//     Term 34 (AT2200-0500)/CC Inputs/Current actual value Ch.23 <-> Data Pointer/CurrentActualValues[22]
//     Term 34 (AT2200-0500)/CC Inputs/Current actual value Ch.24 <-> Data Pointer/CurrentActualValues[23]
//     Term 34 (AT2200-0500)/CC Inputs/Current actual value Ch.25 <-> Data Pointer/CurrentActualValues[24]
//     Term 34 (AT2200-0500)/CC Inputs/Current actual value Ch.26 <-> Data Pointer/CurrentActualValues[25]
//     Term 34 (AT2200-0500)/CC Inputs/Current actual value Ch.27 <-> Data Pointer/CurrentActualValues[26]
//     Term 34 (AT2200-0500)/CC Inputs/Current actual value Ch.28 <-> Data Pointer/CurrentActualValues[27]
//     Term 34 (AT2200-0500)/CC Inputs/Current actual value Ch.29 <-> Data Pointer/CurrentActualValues[28]
//     Term 34 (AT2200-0500)/CC Inputs/Current actual value Ch.3 <-> Data Pointer/CurrentActualValues[2]
//     Term 34 (AT2200-0500)/CC Inputs/Current actual value Ch.30 <-> Data Pointer/CurrentActualValues[29]
//     Term 34 (AT2200-0500)/CC Inputs/Current actual value Ch.4 <-> Data Pointer/CurrentActualValues[3]
//     Term 34 (AT2200-0500)/CC Inputs/Current actual value Ch.5 <-> Data Pointer/CurrentActualValues[4]
//     Term 34 (AT2200-0500)/CC Inputs/Current actual value Ch.6 <-> Data Pointer/CurrentActualValues[5]
//     Term 34 (AT2200-0500)/CC Inputs/Current actual value Ch.7 <-> Data Pointer/CurrentActualValues[6]
//     Term 34 (AT2200-0500)/CC Inputs/Current actual value Ch.8 <-> Data Pointer/CurrentActualValues[7]
//     Term 34 (AT2200-0500)/CC Inputs/Current actual value Ch.9 <-> Data Pointer/CurrentActualValues[8]
//     Term 34 (AT2200-0500)/CC Inputs/Status <-> Data Pointer/Status
//     Term 34 (AT2200-0500)/CC Outputs/Control <-> Data Pointer/Control
//     Term 34 (AT2200-0500)/CC Outputs/Current setpoint value Ch.1 <-> Data Pointer/CurrentSetpointValues[0]
//     Term 34 (AT2200-0500)/CC Outputs/Current setpoint value Ch.10 <-> Data Pointer/CurrentSetpointValues[9]
//     Term 34 (AT2200-0500)/CC Outputs/Current setpoint value Ch.11 <-> Data Pointer/CurrentSetpointValues[10]
//     Term 34 (AT2200-0500)/CC Outputs/Current setpoint value Ch.12 <-> Data Pointer/CurrentSetpointValues[11]
//     Term 34 (AT2200-0500)/CC Outputs/Current setpoint value Ch.13 <-> Data Pointer/CurrentSetpointValues[12]
//     Term 34 (AT2200-0500)/CC Outputs/Current setpoint value Ch.14 <-> Data Pointer/CurrentSetpointValues[13]
//     Term 34 (AT2200-0500)/CC Outputs/Current setpoint value Ch.15 <-> Data Pointer/CurrentSetpointValues[14]
//     Term 34 (AT2200-0500)/CC Outputs/Current setpoint value Ch.16 <-> Data Pointer/CurrentSetpointValues[15]
//     Term 34 (AT2200-0500)/CC Outputs/Current setpoint value Ch.17 <-> Data Pointer/CurrentSetpointValues[16]
//     Term 34 (AT2200-0500)/CC Outputs/Current setpoint value Ch.18 <-> Data Pointer/CurrentSetpointValues[17]
//     Term 34 (AT2200-0500)/CC Outputs/Current setpoint value Ch.19 <-> Data Pointer/CurrentSetpointValues[18]
//     Term 34 (AT2200-0500)/CC Outputs/Current setpoint value Ch.2 <-> Data Pointer/CurrentSetpointValues[1]
//     Term 34 (AT2200-0500)/CC Outputs/Current setpoint value Ch.20 <-> Data Pointer/CurrentSetpointValues[19]
//     Term 34 (AT2200-0500)/CC Outputs/Current setpoint value Ch.21 <-> Data Pointer/CurrentSetpointValues[20]
//     Term 34 (AT2200-0500)/CC Outputs/Current setpoint value Ch.22 <-> Data Pointer/CurrentSetpointValues[21]
//     Term 34 (AT2200-0500)/CC Outputs/Current setpoint value Ch.23 <-> Data Pointer/CurrentSetpointValues[22]
//     Term 34 (AT2200-0500)/CC Outputs/Current setpoint value Ch.24 <-> Data Pointer/CurrentSetpointValues[23]
//     Term 34 (AT2200-0500)/CC Outputs/Current setpoint value Ch.25 <-> Data Pointer/CurrentSetpointValues[24]
//     Term 34 (AT2200-0500)/CC Outputs/Current setpoint value Ch.26 <-> Data Pointer/CurrentSetpointValues[25]
//     Term 34 (AT2200-0500)/CC Outputs/Current setpoint value Ch.27 <-> Data Pointer/CurrentSetpointValues[26]
//     Term 34 (AT2200-0500)/CC Outputs/Current setpoint value Ch.28 <-> Data Pointer/CurrentSetpointValues[27]
//     Term 34 (AT2200-0500)/CC Outputs/Current setpoint value Ch.29 <-> Data Pointer/CurrentSetpointValues[28]
//     Term 34 (AT2200-0500)/CC Outputs/Current setpoint value Ch.3 <-> Data Pointer/CurrentSetpointValues[2]
//     Term 34 (AT2200-0500)/CC Outputs/Current setpoint value Ch.30 <-> Data Pointer/CurrentSetpointValues[29]
//     Term 34 (AT2200-0500)/CC Outputs/Current setpoint value Ch.4 <-> Data Pointer/CurrentSetpointValues[3]
//     Term 34 (AT2200-0500)/CC Outputs/Current setpoint value Ch.5 <-> Data Pointer/CurrentSetpointValues[4]
//     Term 34 (AT2200-0500)/CC Outputs/Current setpoint value Ch.6 <-> Data Pointer/CurrentSetpointValues[5]
//     Term 34 (AT2200-0500)/CC Outputs/Current setpoint value Ch.7 <-> Data Pointer/CurrentSetpointValues[6]
//     Term 34 (AT2200-0500)/CC Outputs/Current setpoint value Ch.8 <-> Data Pointer/CurrentSetpointValues[7]
//     Term 34 (AT2200-0500)/CC Outputs/Current setpoint value Ch.9 <-> Data Pointer/CurrentSetpointValues[8]
//     Term 34 (AT2200-0500)/LFB Inputs/BinaryData <-> Data Pointer/HallSensorValues
//   Device 36 <-> TcCOM Objects/XTS ProcessingUnit 1/Part 1/Module 42
//     Term 35 (AT2200-0500)/CC Inputs/Current actual value Ch.1 <-> Data Pointer/CurrentActualValues[0]
//     Term 35 (AT2200-0500)/CC Inputs/Current actual value Ch.10 <-> Data Pointer/CurrentActualValues[9]
//     Term 35 (AT2200-0500)/CC Inputs/Current actual value Ch.11 <-> Data Pointer/CurrentActualValues[10]
//     Term 35 (AT2200-0500)/CC Inputs/Current actual value Ch.12 <-> Data Pointer/CurrentActualValues[11]
//     Term 35 (AT2200-0500)/CC Inputs/Current actual value Ch.13 <-> Data Pointer/CurrentActualValues[12]
//     Term 35 (AT2200-0500)/CC Inputs/Current actual value Ch.14 <-> Data Pointer/CurrentActualValues[13]
//     Term 35 (AT2200-0500)/CC Inputs/Current actual value Ch.15 <-> Data Pointer/CurrentActualValues[14]
//     Term 35 (AT2200-0500)/CC Inputs/Current actual value Ch.16 <-> Data Pointer/CurrentActualValues[15]
//     Term 35 (AT2200-0500)/CC Inputs/Current actual value Ch.17 <-> Data Pointer/CurrentActualValues[16]
//     Term 35 (AT2200-0500)/CC Inputs/Current actual value Ch.18 <-> Data Pointer/CurrentActualValues[17]
//     Term 35 (AT2200-0500)/CC Inputs/Current actual value Ch.19 <-> Data Pointer/CurrentActualValues[18]
//     Term 35 (AT2200-0500)/CC Inputs/Current actual value Ch.2 <-> Data Pointer/CurrentActualValues[1]
//     Term 35 (AT2200-0500)/CC Inputs/Current actual value Ch.20 <-> Data Pointer/CurrentActualValues[19]
//     Term 35 (AT2200-0500)/CC Inputs/Current actual value Ch.21 <-> Data Pointer/CurrentActualValues[20]
//     Term 35 (AT2200-0500)/CC Inputs/Current actual value Ch.22 <-> Data Pointer/CurrentActualValues[21]
//     Term 35 (AT2200-0500)/CC Inputs/Current actual value Ch.23 <-> Data Pointer/CurrentActualValues[22]
//     Term 35 (AT2200-0500)/CC Inputs/Current actual value Ch.24 <-> Data Pointer/CurrentActualValues[23]
//     Term 35 (AT2200-0500)/CC Inputs/Current actual value Ch.25 <-> Data Pointer/CurrentActualValues[24]
//     Term 35 (AT2200-0500)/CC Inputs/Current actual value Ch.26 <-> Data Pointer/CurrentActualValues[25]
//     Term 35 (AT2200-0500)/CC Inputs/Current actual value Ch.27 <-> Data Pointer/CurrentActualValues[26]
//     Term 35 (AT2200-0500)/CC Inputs/Current actual value Ch.28 <-> Data Pointer/CurrentActualValues[27]
//     Term 35 (AT2200-0500)/CC Inputs/Current actual value Ch.29 <-> Data Pointer/CurrentActualValues[28]
//     Term 35 (AT2200-0500)/CC Inputs/Current actual value Ch.3 <-> Data Pointer/CurrentActualValues[2]
//     Term 35 (AT2200-0500)/CC Inputs/Current actual value Ch.30 <-> Data Pointer/CurrentActualValues[29]
//     Term 35 (AT2200-0500)/CC Inputs/Current actual value Ch.4 <-> Data Pointer/CurrentActualValues[3]
//     Term 35 (AT2200-0500)/CC Inputs/Current actual value Ch.5 <-> Data Pointer/CurrentActualValues[4]
//     Term 35 (AT2200-0500)/CC Inputs/Current actual value Ch.6 <-> Data Pointer/CurrentActualValues[5]
//     Term 35 (AT2200-0500)/CC Inputs/Current actual value Ch.7 <-> Data Pointer/CurrentActualValues[6]
//     Term 35 (AT2200-0500)/CC Inputs/Current actual value Ch.8 <-> Data Pointer/CurrentActualValues[7]
//     Term 35 (AT2200-0500)/CC Inputs/Current actual value Ch.9 <-> Data Pointer/CurrentActualValues[8]
//     Term 35 (AT2200-0500)/CC Inputs/Status <-> Data Pointer/Status
//     Term 35 (AT2200-0500)/CC Outputs/Control <-> Data Pointer/Control
//     Term 35 (AT2200-0500)/CC Outputs/Current setpoint value Ch.1 <-> Data Pointer/CurrentSetpointValues[0]
//     Term 35 (AT2200-0500)/CC Outputs/Current setpoint value Ch.10 <-> Data Pointer/CurrentSetpointValues[9]
//     Term 35 (AT2200-0500)/CC Outputs/Current setpoint value Ch.11 <-> Data Pointer/CurrentSetpointValues[10]
//     Term 35 (AT2200-0500)/CC Outputs/Current setpoint value Ch.12 <-> Data Pointer/CurrentSetpointValues[11]
//     Term 35 (AT2200-0500)/CC Outputs/Current setpoint value Ch.13 <-> Data Pointer/CurrentSetpointValues[12]
//     Term 35 (AT2200-0500)/CC Outputs/Current setpoint value Ch.14 <-> Data Pointer/CurrentSetpointValues[13]
//     Term 35 (AT2200-0500)/CC Outputs/Current setpoint value Ch.15 <-> Data Pointer/CurrentSetpointValues[14]
//     Term 35 (AT2200-0500)/CC Outputs/Current setpoint value Ch.16 <-> Data Pointer/CurrentSetpointValues[15]
//     Term 35 (AT2200-0500)/CC Outputs/Current setpoint value Ch.17 <-> Data Pointer/CurrentSetpointValues[16]
//     Term 35 (AT2200-0500)/CC Outputs/Current setpoint value Ch.18 <-> Data Pointer/CurrentSetpointValues[17]
//     Term 35 (AT2200-0500)/CC Outputs/Current setpoint value Ch.19 <-> Data Pointer/CurrentSetpointValues[18]
//     Term 35 (AT2200-0500)/CC Outputs/Current setpoint value Ch.2 <-> Data Pointer/CurrentSetpointValues[1]
//     Term 35 (AT2200-0500)/CC Outputs/Current setpoint value Ch.20 <-> Data Pointer/CurrentSetpointValues[19]
//     Term 35 (AT2200-0500)/CC Outputs/Current setpoint value Ch.21 <-> Data Pointer/CurrentSetpointValues[20]
//     Term 35 (AT2200-0500)/CC Outputs/Current setpoint value Ch.22 <-> Data Pointer/CurrentSetpointValues[21]
//     Term 35 (AT2200-0500)/CC Outputs/Current setpoint value Ch.23 <-> Data Pointer/CurrentSetpointValues[22]
//     Term 35 (AT2200-0500)/CC Outputs/Current setpoint value Ch.24 <-> Data Pointer/CurrentSetpointValues[23]
//     Term 35 (AT2200-0500)/CC Outputs/Current setpoint value Ch.25 <-> Data Pointer/CurrentSetpointValues[24]
//     Term 35 (AT2200-0500)/CC Outputs/Current setpoint value Ch.26 <-> Data Pointer/CurrentSetpointValues[25]
//     Term 35 (AT2200-0500)/CC Outputs/Current setpoint value Ch.27 <-> Data Pointer/CurrentSetpointValues[26]
//     Term 35 (AT2200-0500)/CC Outputs/Current setpoint value Ch.28 <-> Data Pointer/CurrentSetpointValues[27]
//     Term 35 (AT2200-0500)/CC Outputs/Current setpoint value Ch.29 <-> Data Pointer/CurrentSetpointValues[28]
//     Term 35 (AT2200-0500)/CC Outputs/Current setpoint value Ch.3 <-> Data Pointer/CurrentSetpointValues[2]
//     Term 35 (AT2200-0500)/CC Outputs/Current setpoint value Ch.30 <-> Data Pointer/CurrentSetpointValues[29]
//     Term 35 (AT2200-0500)/CC Outputs/Current setpoint value Ch.4 <-> Data Pointer/CurrentSetpointValues[3]
//     Term 35 (AT2200-0500)/CC Outputs/Current setpoint value Ch.5 <-> Data Pointer/CurrentSetpointValues[4]
//     Term 35 (AT2200-0500)/CC Outputs/Current setpoint value Ch.6 <-> Data Pointer/CurrentSetpointValues[5]
//     Term 35 (AT2200-0500)/CC Outputs/Current setpoint value Ch.7 <-> Data Pointer/CurrentSetpointValues[6]
//     Term 35 (AT2200-0500)/CC Outputs/Current setpoint value Ch.8 <-> Data Pointer/CurrentSetpointValues[7]
//     Term 35 (AT2200-0500)/CC Outputs/Current setpoint value Ch.9 <-> Data Pointer/CurrentSetpointValues[8]
//     Term 35 (AT2200-0500)/LFB Inputs/BinaryData <-> Data Pointer/HallSensorValues
//   Device 37 <-> TcCOM Objects/XTS ProcessingUnit 1/Part 1/Module 43
//     Term 36 (AT2202-0500)/CC Inputs/Current actual value Ch.1 <-> Data Pointer/CurrentActualValues[0]
//     Term 36 (AT2202-0500)/CC Inputs/Current actual value Ch.10 <-> Data Pointer/CurrentActualValues[9]
//     Term 36 (AT2202-0500)/CC Inputs/Current actual value Ch.11 <-> Data Pointer/CurrentActualValues[10]
//     Term 36 (AT2202-0500)/CC Inputs/Current actual value Ch.12 <-> Data Pointer/CurrentActualValues[11]
//     Term 36 (AT2202-0500)/CC Inputs/Current actual value Ch.13 <-> Data Pointer/CurrentActualValues[12]
//     Term 36 (AT2202-0500)/CC Inputs/Current actual value Ch.14 <-> Data Pointer/CurrentActualValues[13]
//     Term 36 (AT2202-0500)/CC Inputs/Current actual value Ch.15 <-> Data Pointer/CurrentActualValues[14]
//     Term 36 (AT2202-0500)/CC Inputs/Current actual value Ch.16 <-> Data Pointer/CurrentActualValues[15]
//     Term 36 (AT2202-0500)/CC Inputs/Current actual value Ch.17 <-> Data Pointer/CurrentActualValues[16]
//     Term 36 (AT2202-0500)/CC Inputs/Current actual value Ch.18 <-> Data Pointer/CurrentActualValues[17]
//     Term 36 (AT2202-0500)/CC Inputs/Current actual value Ch.19 <-> Data Pointer/CurrentActualValues[18]
//     Term 36 (AT2202-0500)/CC Inputs/Current actual value Ch.2 <-> Data Pointer/CurrentActualValues[1]
//     Term 36 (AT2202-0500)/CC Inputs/Current actual value Ch.20 <-> Data Pointer/CurrentActualValues[19]
//     Term 36 (AT2202-0500)/CC Inputs/Current actual value Ch.21 <-> Data Pointer/CurrentActualValues[20]
//     Term 36 (AT2202-0500)/CC Inputs/Current actual value Ch.22 <-> Data Pointer/CurrentActualValues[21]
//     Term 36 (AT2202-0500)/CC Inputs/Current actual value Ch.23 <-> Data Pointer/CurrentActualValues[22]
//     Term 36 (AT2202-0500)/CC Inputs/Current actual value Ch.24 <-> Data Pointer/CurrentActualValues[23]
//     Term 36 (AT2202-0500)/CC Inputs/Current actual value Ch.25 <-> Data Pointer/CurrentActualValues[24]
//     Term 36 (AT2202-0500)/CC Inputs/Current actual value Ch.26 <-> Data Pointer/CurrentActualValues[25]
//     Term 36 (AT2202-0500)/CC Inputs/Current actual value Ch.27 <-> Data Pointer/CurrentActualValues[26]
//     Term 36 (AT2202-0500)/CC Inputs/Current actual value Ch.28 <-> Data Pointer/CurrentActualValues[27]
//     Term 36 (AT2202-0500)/CC Inputs/Current actual value Ch.29 <-> Data Pointer/CurrentActualValues[28]
//     Term 36 (AT2202-0500)/CC Inputs/Current actual value Ch.3 <-> Data Pointer/CurrentActualValues[2]
//     Term 36 (AT2202-0500)/CC Inputs/Current actual value Ch.30 <-> Data Pointer/CurrentActualValues[29]
//     Term 36 (AT2202-0500)/CC Inputs/Current actual value Ch.4 <-> Data Pointer/CurrentActualValues[3]
//     Term 36 (AT2202-0500)/CC Inputs/Current actual value Ch.5 <-> Data Pointer/CurrentActualValues[4]
//     Term 36 (AT2202-0500)/CC Inputs/Current actual value Ch.6 <-> Data Pointer/CurrentActualValues[5]
//     Term 36 (AT2202-0500)/CC Inputs/Current actual value Ch.7 <-> Data Pointer/CurrentActualValues[6]
//     Term 36 (AT2202-0500)/CC Inputs/Current actual value Ch.8 <-> Data Pointer/CurrentActualValues[7]
//     Term 36 (AT2202-0500)/CC Inputs/Current actual value Ch.9 <-> Data Pointer/CurrentActualValues[8]
//     Term 36 (AT2202-0500)/CC Inputs/Status <-> Data Pointer/Status
//     Term 36 (AT2202-0500)/CC Outputs/Control <-> Data Pointer/Control
//     Term 36 (AT2202-0500)/CC Outputs/Current setpoint value Ch.1 <-> Data Pointer/CurrentSetpointValues[0]
//     Term 36 (AT2202-0500)/CC Outputs/Current setpoint value Ch.10 <-> Data Pointer/CurrentSetpointValues[9]
//     Term 36 (AT2202-0500)/CC Outputs/Current setpoint value Ch.11 <-> Data Pointer/CurrentSetpointValues[10]
//     Term 36 (AT2202-0500)/CC Outputs/Current setpoint value Ch.12 <-> Data Pointer/CurrentSetpointValues[11]
//     Term 36 (AT2202-0500)/CC Outputs/Current setpoint value Ch.13 <-> Data Pointer/CurrentSetpointValues[12]
//     Term 36 (AT2202-0500)/CC Outputs/Current setpoint value Ch.14 <-> Data Pointer/CurrentSetpointValues[13]
//     Term 36 (AT2202-0500)/CC Outputs/Current setpoint value Ch.15 <-> Data Pointer/CurrentSetpointValues[14]
//     Term 36 (AT2202-0500)/CC Outputs/Current setpoint value Ch.16 <-> Data Pointer/CurrentSetpointValues[15]
//     Term 36 (AT2202-0500)/CC Outputs/Current setpoint value Ch.17 <-> Data Pointer/CurrentSetpointValues[16]
//     Term 36 (AT2202-0500)/CC Outputs/Current setpoint value Ch.18 <-> Data Pointer/CurrentSetpointValues[17]
//     Term 36 (AT2202-0500)/CC Outputs/Current setpoint value Ch.19 <-> Data Pointer/CurrentSetpointValues[18]
//     Term 36 (AT2202-0500)/CC Outputs/Current setpoint value Ch.2 <-> Data Pointer/CurrentSetpointValues[1]
//     Term 36 (AT2202-0500)/CC Outputs/Current setpoint value Ch.20 <-> Data Pointer/CurrentSetpointValues[19]
//     Term 36 (AT2202-0500)/CC Outputs/Current setpoint value Ch.21 <-> Data Pointer/CurrentSetpointValues[20]
//     Term 36 (AT2202-0500)/CC Outputs/Current setpoint value Ch.22 <-> Data Pointer/CurrentSetpointValues[21]
//     Term 36 (AT2202-0500)/CC Outputs/Current setpoint value Ch.23 <-> Data Pointer/CurrentSetpointValues[22]
//     Term 36 (AT2202-0500)/CC Outputs/Current setpoint value Ch.24 <-> Data Pointer/CurrentSetpointValues[23]
//     Term 36 (AT2202-0500)/CC Outputs/Current setpoint value Ch.25 <-> Data Pointer/CurrentSetpointValues[24]
//     Term 36 (AT2202-0500)/CC Outputs/Current setpoint value Ch.26 <-> Data Pointer/CurrentSetpointValues[25]
//     Term 36 (AT2202-0500)/CC Outputs/Current setpoint value Ch.27 <-> Data Pointer/CurrentSetpointValues[26]
//     Term 36 (AT2202-0500)/CC Outputs/Current setpoint value Ch.28 <-> Data Pointer/CurrentSetpointValues[27]
//     Term 36 (AT2202-0500)/CC Outputs/Current setpoint value Ch.29 <-> Data Pointer/CurrentSetpointValues[28]
//     Term 36 (AT2202-0500)/CC Outputs/Current setpoint value Ch.3 <-> Data Pointer/CurrentSetpointValues[2]
//     Term 36 (AT2202-0500)/CC Outputs/Current setpoint value Ch.30 <-> Data Pointer/CurrentSetpointValues[29]
//     Term 36 (AT2202-0500)/CC Outputs/Current setpoint value Ch.4 <-> Data Pointer/CurrentSetpointValues[3]
//     Term 36 (AT2202-0500)/CC Outputs/Current setpoint value Ch.5 <-> Data Pointer/CurrentSetpointValues[4]
//     Term 36 (AT2202-0500)/CC Outputs/Current setpoint value Ch.6 <-> Data Pointer/CurrentSetpointValues[5]
//     Term 36 (AT2202-0500)/CC Outputs/Current setpoint value Ch.7 <-> Data Pointer/CurrentSetpointValues[6]
//     Term 36 (AT2202-0500)/CC Outputs/Current setpoint value Ch.8 <-> Data Pointer/CurrentSetpointValues[7]
//     Term 36 (AT2202-0500)/CC Outputs/Current setpoint value Ch.9 <-> Data Pointer/CurrentSetpointValues[8]
//     Term 36 (AT2202-0500)/LFB Inputs/BinaryData <-> Data Pointer/HallSensorValues
//   Device 37 <-> TcCOM Objects/XTS ProcessingUnit 1/Part 1/Module 44
//     Term 37 (AT2200-0500)/CC Inputs/Current actual value Ch.1 <-> Data Pointer/CurrentActualValues[0]
//     Term 37 (AT2200-0500)/CC Inputs/Current actual value Ch.10 <-> Data Pointer/CurrentActualValues[9]
//     Term 37 (AT2200-0500)/CC Inputs/Current actual value Ch.11 <-> Data Pointer/CurrentActualValues[10]
//     Term 37 (AT2200-0500)/CC Inputs/Current actual value Ch.12 <-> Data Pointer/CurrentActualValues[11]
//     Term 37 (AT2200-0500)/CC Inputs/Current actual value Ch.13 <-> Data Pointer/CurrentActualValues[12]
//     Term 37 (AT2200-0500)/CC Inputs/Current actual value Ch.14 <-> Data Pointer/CurrentActualValues[13]
//     Term 37 (AT2200-0500)/CC Inputs/Current actual value Ch.15 <-> Data Pointer/CurrentActualValues[14]
//     Term 37 (AT2200-0500)/CC Inputs/Current actual value Ch.16 <-> Data Pointer/CurrentActualValues[15]
//     Term 37 (AT2200-0500)/CC Inputs/Current actual value Ch.17 <-> Data Pointer/CurrentActualValues[16]
//     Term 37 (AT2200-0500)/CC Inputs/Current actual value Ch.18 <-> Data Pointer/CurrentActualValues[17]
//     Term 37 (AT2200-0500)/CC Inputs/Current actual value Ch.19 <-> Data Pointer/CurrentActualValues[18]
//     Term 37 (AT2200-0500)/CC Inputs/Current actual value Ch.2 <-> Data Pointer/CurrentActualValues[1]
//     Term 37 (AT2200-0500)/CC Inputs/Current actual value Ch.20 <-> Data Pointer/CurrentActualValues[19]
//     Term 37 (AT2200-0500)/CC Inputs/Current actual value Ch.21 <-> Data Pointer/CurrentActualValues[20]
//     Term 37 (AT2200-0500)/CC Inputs/Current actual value Ch.22 <-> Data Pointer/CurrentActualValues[21]
//     Term 37 (AT2200-0500)/CC Inputs/Current actual value Ch.23 <-> Data Pointer/CurrentActualValues[22]
//     Term 37 (AT2200-0500)/CC Inputs/Current actual value Ch.24 <-> Data Pointer/CurrentActualValues[23]
//     Term 37 (AT2200-0500)/CC Inputs/Current actual value Ch.25 <-> Data Pointer/CurrentActualValues[24]
//     Term 37 (AT2200-0500)/CC Inputs/Current actual value Ch.26 <-> Data Pointer/CurrentActualValues[25]
//     Term 37 (AT2200-0500)/CC Inputs/Current actual value Ch.27 <-> Data Pointer/CurrentActualValues[26]
//     Term 37 (AT2200-0500)/CC Inputs/Current actual value Ch.28 <-> Data Pointer/CurrentActualValues[27]
//     Term 37 (AT2200-0500)/CC Inputs/Current actual value Ch.29 <-> Data Pointer/CurrentActualValues[28]
//     Term 37 (AT2200-0500)/CC Inputs/Current actual value Ch.3 <-> Data Pointer/CurrentActualValues[2]
//     Term 37 (AT2200-0500)/CC Inputs/Current actual value Ch.30 <-> Data Pointer/CurrentActualValues[29]
//     Term 37 (AT2200-0500)/CC Inputs/Current actual value Ch.4 <-> Data Pointer/CurrentActualValues[3]
//     Term 37 (AT2200-0500)/CC Inputs/Current actual value Ch.5 <-> Data Pointer/CurrentActualValues[4]
//     Term 37 (AT2200-0500)/CC Inputs/Current actual value Ch.6 <-> Data Pointer/CurrentActualValues[5]
//     Term 37 (AT2200-0500)/CC Inputs/Current actual value Ch.7 <-> Data Pointer/CurrentActualValues[6]
//     Term 37 (AT2200-0500)/CC Inputs/Current actual value Ch.8 <-> Data Pointer/CurrentActualValues[7]
//     Term 37 (AT2200-0500)/CC Inputs/Current actual value Ch.9 <-> Data Pointer/CurrentActualValues[8]
//     Term 37 (AT2200-0500)/CC Inputs/Status <-> Data Pointer/Status
//     Term 37 (AT2200-0500)/CC Outputs/Control <-> Data Pointer/Control
//     Term 37 (AT2200-0500)/CC Outputs/Current setpoint value Ch.1 <-> Data Pointer/CurrentSetpointValues[0]
//     Term 37 (AT2200-0500)/CC Outputs/Current setpoint value Ch.10 <-> Data Pointer/CurrentSetpointValues[9]
//     Term 37 (AT2200-0500)/CC Outputs/Current setpoint value Ch.11 <-> Data Pointer/CurrentSetpointValues[10]
//     Term 37 (AT2200-0500)/CC Outputs/Current setpoint value Ch.12 <-> Data Pointer/CurrentSetpointValues[11]
//     Term 37 (AT2200-0500)/CC Outputs/Current setpoint value Ch.13 <-> Data Pointer/CurrentSetpointValues[12]
//     Term 37 (AT2200-0500)/CC Outputs/Current setpoint value Ch.14 <-> Data Pointer/CurrentSetpointValues[13]
//     Term 37 (AT2200-0500)/CC Outputs/Current setpoint value Ch.15 <-> Data Pointer/CurrentSetpointValues[14]
//     Term 37 (AT2200-0500)/CC Outputs/Current setpoint value Ch.16 <-> Data Pointer/CurrentSetpointValues[15]
//     Term 37 (AT2200-0500)/CC Outputs/Current setpoint value Ch.17 <-> Data Pointer/CurrentSetpointValues[16]
//     Term 37 (AT2200-0500)/CC Outputs/Current setpoint value Ch.18 <-> Data Pointer/CurrentSetpointValues[17]
//     Term 37 (AT2200-0500)/CC Outputs/Current setpoint value Ch.19 <-> Data Pointer/CurrentSetpointValues[18]
//     Term 37 (AT2200-0500)/CC Outputs/Current setpoint value Ch.2 <-> Data Pointer/CurrentSetpointValues[1]
//     Term 37 (AT2200-0500)/CC Outputs/Current setpoint value Ch.20 <-> Data Pointer/CurrentSetpointValues[19]
//     Term 37 (AT2200-0500)/CC Outputs/Current setpoint value Ch.21 <-> Data Pointer/CurrentSetpointValues[20]
//     Term 37 (AT2200-0500)/CC Outputs/Current setpoint value Ch.22 <-> Data Pointer/CurrentSetpointValues[21]
//     Term 37 (AT2200-0500)/CC Outputs/Current setpoint value Ch.23 <-> Data Pointer/CurrentSetpointValues[22]
//     Term 37 (AT2200-0500)/CC Outputs/Current setpoint value Ch.24 <-> Data Pointer/CurrentSetpointValues[23]
//     Term 37 (AT2200-0500)/CC Outputs/Current setpoint value Ch.25 <-> Data Pointer/CurrentSetpointValues[24]
//     Term 37 (AT2200-0500)/CC Outputs/Current setpoint value Ch.26 <-> Data Pointer/CurrentSetpointValues[25]
//     Term 37 (AT2200-0500)/CC Outputs/Current setpoint value Ch.27 <-> Data Pointer/CurrentSetpointValues[26]
//     Term 37 (AT2200-0500)/CC Outputs/Current setpoint value Ch.28 <-> Data Pointer/CurrentSetpointValues[27]
//     Term 37 (AT2200-0500)/CC Outputs/Current setpoint value Ch.29 <-> Data Pointer/CurrentSetpointValues[28]
//     Term 37 (AT2200-0500)/CC Outputs/Current setpoint value Ch.3 <-> Data Pointer/CurrentSetpointValues[2]
//     Term 37 (AT2200-0500)/CC Outputs/Current setpoint value Ch.30 <-> Data Pointer/CurrentSetpointValues[29]
//     Term 37 (AT2200-0500)/CC Outputs/Current setpoint value Ch.4 <-> Data Pointer/CurrentSetpointValues[3]
//     Term 37 (AT2200-0500)/CC Outputs/Current setpoint value Ch.5 <-> Data Pointer/CurrentSetpointValues[4]
//     Term 37 (AT2200-0500)/CC Outputs/Current setpoint value Ch.6 <-> Data Pointer/CurrentSetpointValues[5]
//     Term 37 (AT2200-0500)/CC Outputs/Current setpoint value Ch.7 <-> Data Pointer/CurrentSetpointValues[6]
//     Term 37 (AT2200-0500)/CC Outputs/Current setpoint value Ch.8 <-> Data Pointer/CurrentSetpointValues[7]
//     Term 37 (AT2200-0500)/CC Outputs/Current setpoint value Ch.9 <-> Data Pointer/CurrentSetpointValues[8]
//     Term 37 (AT2200-0500)/LFB Inputs/BinaryData <-> Data Pointer/HallSensorValues
//   Device 37 <-> TcCOM Objects/XTS ProcessingUnit 1/Part 1/Module 45
//     Term 38 (AT2200-0500)/CC Inputs/Current actual value Ch.1 <-> Data Pointer/CurrentActualValues[0]
//     Term 38 (AT2200-0500)/CC Inputs/Current actual value Ch.10 <-> Data Pointer/CurrentActualValues[9]
//     Term 38 (AT2200-0500)/CC Inputs/Current actual value Ch.11 <-> Data Pointer/CurrentActualValues[10]
//     Term 38 (AT2200-0500)/CC Inputs/Current actual value Ch.12 <-> Data Pointer/CurrentActualValues[11]
//     Term 38 (AT2200-0500)/CC Inputs/Current actual value Ch.13 <-> Data Pointer/CurrentActualValues[12]
//     Term 38 (AT2200-0500)/CC Inputs/Current actual value Ch.14 <-> Data Pointer/CurrentActualValues[13]
//     Term 38 (AT2200-0500)/CC Inputs/Current actual value Ch.15 <-> Data Pointer/CurrentActualValues[14]
//     Term 38 (AT2200-0500)/CC Inputs/Current actual value Ch.16 <-> Data Pointer/CurrentActualValues[15]
//     Term 38 (AT2200-0500)/CC Inputs/Current actual value Ch.17 <-> Data Pointer/CurrentActualValues[16]
//     Term 38 (AT2200-0500)/CC Inputs/Current actual value Ch.18 <-> Data Pointer/CurrentActualValues[17]
//     Term 38 (AT2200-0500)/CC Inputs/Current actual value Ch.19 <-> Data Pointer/CurrentActualValues[18]
//     Term 38 (AT2200-0500)/CC Inputs/Current actual value Ch.2 <-> Data Pointer/CurrentActualValues[1]
//     Term 38 (AT2200-0500)/CC Inputs/Current actual value Ch.20 <-> Data Pointer/CurrentActualValues[19]
//     Term 38 (AT2200-0500)/CC Inputs/Current actual value Ch.21 <-> Data Pointer/CurrentActualValues[20]
//     Term 38 (AT2200-0500)/CC Inputs/Current actual value Ch.22 <-> Data Pointer/CurrentActualValues[21]
//     Term 38 (AT2200-0500)/CC Inputs/Current actual value Ch.23 <-> Data Pointer/CurrentActualValues[22]
//     Term 38 (AT2200-0500)/CC Inputs/Current actual value Ch.24 <-> Data Pointer/CurrentActualValues[23]
//     Term 38 (AT2200-0500)/CC Inputs/Current actual value Ch.25 <-> Data Pointer/CurrentActualValues[24]
//     Term 38 (AT2200-0500)/CC Inputs/Current actual value Ch.26 <-> Data Pointer/CurrentActualValues[25]
//     Term 38 (AT2200-0500)/CC Inputs/Current actual value Ch.27 <-> Data Pointer/CurrentActualValues[26]
//     Term 38 (AT2200-0500)/CC Inputs/Current actual value Ch.28 <-> Data Pointer/CurrentActualValues[27]
//     Term 38 (AT2200-0500)/CC Inputs/Current actual value Ch.29 <-> Data Pointer/CurrentActualValues[28]
//     Term 38 (AT2200-0500)/CC Inputs/Current actual value Ch.3 <-> Data Pointer/CurrentActualValues[2]
//     Term 38 (AT2200-0500)/CC Inputs/Current actual value Ch.30 <-> Data Pointer/CurrentActualValues[29]
//     Term 38 (AT2200-0500)/CC Inputs/Current actual value Ch.4 <-> Data Pointer/CurrentActualValues[3]
//     Term 38 (AT2200-0500)/CC Inputs/Current actual value Ch.5 <-> Data Pointer/CurrentActualValues[4]
//     Term 38 (AT2200-0500)/CC Inputs/Current actual value Ch.6 <-> Data Pointer/CurrentActualValues[5]
//     Term 38 (AT2200-0500)/CC Inputs/Current actual value Ch.7 <-> Data Pointer/CurrentActualValues[6]
//     Term 38 (AT2200-0500)/CC Inputs/Current actual value Ch.8 <-> Data Pointer/CurrentActualValues[7]
//     Term 38 (AT2200-0500)/CC Inputs/Current actual value Ch.9 <-> Data Pointer/CurrentActualValues[8]
//     Term 38 (AT2200-0500)/CC Inputs/Status <-> Data Pointer/Status
//     Term 38 (AT2200-0500)/CC Outputs/Control <-> Data Pointer/Control
//     Term 38 (AT2200-0500)/CC Outputs/Current setpoint value Ch.1 <-> Data Pointer/CurrentSetpointValues[0]
//     Term 38 (AT2200-0500)/CC Outputs/Current setpoint value Ch.10 <-> Data Pointer/CurrentSetpointValues[9]
//     Term 38 (AT2200-0500)/CC Outputs/Current setpoint value Ch.11 <-> Data Pointer/CurrentSetpointValues[10]
//     Term 38 (AT2200-0500)/CC Outputs/Current setpoint value Ch.12 <-> Data Pointer/CurrentSetpointValues[11]
//     Term 38 (AT2200-0500)/CC Outputs/Current setpoint value Ch.13 <-> Data Pointer/CurrentSetpointValues[12]
//     Term 38 (AT2200-0500)/CC Outputs/Current setpoint value Ch.14 <-> Data Pointer/CurrentSetpointValues[13]
//     Term 38 (AT2200-0500)/CC Outputs/Current setpoint value Ch.15 <-> Data Pointer/CurrentSetpointValues[14]
//     Term 38 (AT2200-0500)/CC Outputs/Current setpoint value Ch.16 <-> Data Pointer/CurrentSetpointValues[15]
//     Term 38 (AT2200-0500)/CC Outputs/Current setpoint value Ch.17 <-> Data Pointer/CurrentSetpointValues[16]
//     Term 38 (AT2200-0500)/CC Outputs/Current setpoint value Ch.18 <-> Data Pointer/CurrentSetpointValues[17]
//     Term 38 (AT2200-0500)/CC Outputs/Current setpoint value Ch.19 <-> Data Pointer/CurrentSetpointValues[18]
//     Term 38 (AT2200-0500)/CC Outputs/Current setpoint value Ch.2 <-> Data Pointer/CurrentSetpointValues[1]
//     Term 38 (AT2200-0500)/CC Outputs/Current setpoint value Ch.20 <-> Data Pointer/CurrentSetpointValues[19]
//     Term 38 (AT2200-0500)/CC Outputs/Current setpoint value Ch.21 <-> Data Pointer/CurrentSetpointValues[20]
//     Term 38 (AT2200-0500)/CC Outputs/Current setpoint value Ch.22 <-> Data Pointer/CurrentSetpointValues[21]
//     Term 38 (AT2200-0500)/CC Outputs/Current setpoint value Ch.23 <-> Data Pointer/CurrentSetpointValues[22]
//     Term 38 (AT2200-0500)/CC Outputs/Current setpoint value Ch.24 <-> Data Pointer/CurrentSetpointValues[23]
//     Term 38 (AT2200-0500)/CC Outputs/Current setpoint value Ch.25 <-> Data Pointer/CurrentSetpointValues[24]
//     Term 38 (AT2200-0500)/CC Outputs/Current setpoint value Ch.26 <-> Data Pointer/CurrentSetpointValues[25]
//     Term 38 (AT2200-0500)/CC Outputs/Current setpoint value Ch.27 <-> Data Pointer/CurrentSetpointValues[26]
//     Term 38 (AT2200-0500)/CC Outputs/Current setpoint value Ch.28 <-> Data Pointer/CurrentSetpointValues[27]
//     Term 38 (AT2200-0500)/CC Outputs/Current setpoint value Ch.29 <-> Data Pointer/CurrentSetpointValues[28]
//     Term 38 (AT2200-0500)/CC Outputs/Current setpoint value Ch.3 <-> Data Pointer/CurrentSetpointValues[2]
//     Term 38 (AT2200-0500)/CC Outputs/Current setpoint value Ch.30 <-> Data Pointer/CurrentSetpointValues[29]
//     Term 38 (AT2200-0500)/CC Outputs/Current setpoint value Ch.4 <-> Data Pointer/CurrentSetpointValues[3]
//     Term 38 (AT2200-0500)/CC Outputs/Current setpoint value Ch.5 <-> Data Pointer/CurrentSetpointValues[4]
//     Term 38 (AT2200-0500)/CC Outputs/Current setpoint value Ch.6 <-> Data Pointer/CurrentSetpointValues[5]
//     Term 38 (AT2200-0500)/CC Outputs/Current setpoint value Ch.7 <-> Data Pointer/CurrentSetpointValues[6]
//     Term 38 (AT2200-0500)/CC Outputs/Current setpoint value Ch.8 <-> Data Pointer/CurrentSetpointValues[7]
//     Term 38 (AT2200-0500)/CC Outputs/Current setpoint value Ch.9 <-> Data Pointer/CurrentSetpointValues[8]
//     Term 38 (AT2200-0500)/LFB Inputs/BinaryData <-> Data Pointer/HallSensorValues
//   Device 38 <-> TcCOM Objects/XTS ProcessingUnit 1/Part 1/Module 46
//     Term 39 (AT2202-0500)/CC Inputs/Current actual value Ch.1 <-> Data Pointer/CurrentActualValues[0]
//     Term 39 (AT2202-0500)/CC Inputs/Current actual value Ch.10 <-> Data Pointer/CurrentActualValues[9]
//     Term 39 (AT2202-0500)/CC Inputs/Current actual value Ch.11 <-> Data Pointer/CurrentActualValues[10]
//     Term 39 (AT2202-0500)/CC Inputs/Current actual value Ch.12 <-> Data Pointer/CurrentActualValues[11]
//     Term 39 (AT2202-0500)/CC Inputs/Current actual value Ch.13 <-> Data Pointer/CurrentActualValues[12]
//     Term 39 (AT2202-0500)/CC Inputs/Current actual value Ch.14 <-> Data Pointer/CurrentActualValues[13]
//     Term 39 (AT2202-0500)/CC Inputs/Current actual value Ch.15 <-> Data Pointer/CurrentActualValues[14]
//     Term 39 (AT2202-0500)/CC Inputs/Current actual value Ch.16 <-> Data Pointer/CurrentActualValues[15]
//     Term 39 (AT2202-0500)/CC Inputs/Current actual value Ch.17 <-> Data Pointer/CurrentActualValues[16]
//     Term 39 (AT2202-0500)/CC Inputs/Current actual value Ch.18 <-> Data Pointer/CurrentActualValues[17]
//     Term 39 (AT2202-0500)/CC Inputs/Current actual value Ch.19 <-> Data Pointer/CurrentActualValues[18]
//     Term 39 (AT2202-0500)/CC Inputs/Current actual value Ch.2 <-> Data Pointer/CurrentActualValues[1]
//     Term 39 (AT2202-0500)/CC Inputs/Current actual value Ch.20 <-> Data Pointer/CurrentActualValues[19]
//     Term 39 (AT2202-0500)/CC Inputs/Current actual value Ch.21 <-> Data Pointer/CurrentActualValues[20]
//     Term 39 (AT2202-0500)/CC Inputs/Current actual value Ch.22 <-> Data Pointer/CurrentActualValues[21]
//     Term 39 (AT2202-0500)/CC Inputs/Current actual value Ch.23 <-> Data Pointer/CurrentActualValues[22]
//     Term 39 (AT2202-0500)/CC Inputs/Current actual value Ch.24 <-> Data Pointer/CurrentActualValues[23]
//     Term 39 (AT2202-0500)/CC Inputs/Current actual value Ch.25 <-> Data Pointer/CurrentActualValues[24]
//     Term 39 (AT2202-0500)/CC Inputs/Current actual value Ch.26 <-> Data Pointer/CurrentActualValues[25]
//     Term 39 (AT2202-0500)/CC Inputs/Current actual value Ch.27 <-> Data Pointer/CurrentActualValues[26]
//     Term 39 (AT2202-0500)/CC Inputs/Current actual value Ch.28 <-> Data Pointer/CurrentActualValues[27]
//     Term 39 (AT2202-0500)/CC Inputs/Current actual value Ch.29 <-> Data Pointer/CurrentActualValues[28]
//     Term 39 (AT2202-0500)/CC Inputs/Current actual value Ch.3 <-> Data Pointer/CurrentActualValues[2]
//     Term 39 (AT2202-0500)/CC Inputs/Current actual value Ch.30 <-> Data Pointer/CurrentActualValues[29]
//     Term 39 (AT2202-0500)/CC Inputs/Current actual value Ch.4 <-> Data Pointer/CurrentActualValues[3]
//     Term 39 (AT2202-0500)/CC Inputs/Current actual value Ch.5 <-> Data Pointer/CurrentActualValues[4]
//     Term 39 (AT2202-0500)/CC Inputs/Current actual value Ch.6 <-> Data Pointer/CurrentActualValues[5]
//     Term 39 (AT2202-0500)/CC Inputs/Current actual value Ch.7 <-> Data Pointer/CurrentActualValues[6]
//     Term 39 (AT2202-0500)/CC Inputs/Current actual value Ch.8 <-> Data Pointer/CurrentActualValues[7]
//     Term 39 (AT2202-0500)/CC Inputs/Current actual value Ch.9 <-> Data Pointer/CurrentActualValues[8]
//     Term 39 (AT2202-0500)/CC Inputs/Status <-> Data Pointer/Status
//     Term 39 (AT2202-0500)/CC Outputs/Control <-> Data Pointer/Control
//     Term 39 (AT2202-0500)/CC Outputs/Current setpoint value Ch.1 <-> Data Pointer/CurrentSetpointValues[0]
//     Term 39 (AT2202-0500)/CC Outputs/Current setpoint value Ch.10 <-> Data Pointer/CurrentSetpointValues[9]
//     Term 39 (AT2202-0500)/CC Outputs/Current setpoint value Ch.11 <-> Data Pointer/CurrentSetpointValues[10]
//     Term 39 (AT2202-0500)/CC Outputs/Current setpoint value Ch.12 <-> Data Pointer/CurrentSetpointValues[11]
//     Term 39 (AT2202-0500)/CC Outputs/Current setpoint value Ch.13 <-> Data Pointer/CurrentSetpointValues[12]
//     Term 39 (AT2202-0500)/CC Outputs/Current setpoint value Ch.14 <-> Data Pointer/CurrentSetpointValues[13]
//     Term 39 (AT2202-0500)/CC Outputs/Current setpoint value Ch.15 <-> Data Pointer/CurrentSetpointValues[14]
//     Term 39 (AT2202-0500)/CC Outputs/Current setpoint value Ch.16 <-> Data Pointer/CurrentSetpointValues[15]
//     Term 39 (AT2202-0500)/CC Outputs/Current setpoint value Ch.17 <-> Data Pointer/CurrentSetpointValues[16]
//     Term 39 (AT2202-0500)/CC Outputs/Current setpoint value Ch.18 <-> Data Pointer/CurrentSetpointValues[17]
//     Term 39 (AT2202-0500)/CC Outputs/Current setpoint value Ch.19 <-> Data Pointer/CurrentSetpointValues[18]
//     Term 39 (AT2202-0500)/CC Outputs/Current setpoint value Ch.2 <-> Data Pointer/CurrentSetpointValues[1]
//     Term 39 (AT2202-0500)/CC Outputs/Current setpoint value Ch.20 <-> Data Pointer/CurrentSetpointValues[19]
//     Term 39 (AT2202-0500)/CC Outputs/Current setpoint value Ch.21 <-> Data Pointer/CurrentSetpointValues[20]
//     Term 39 (AT2202-0500)/CC Outputs/Current setpoint value Ch.22 <-> Data Pointer/CurrentSetpointValues[21]
//     Term 39 (AT2202-0500)/CC Outputs/Current setpoint value Ch.23 <-> Data Pointer/CurrentSetpointValues[22]
//     Term 39 (AT2202-0500)/CC Outputs/Current setpoint value Ch.24 <-> Data Pointer/CurrentSetpointValues[23]
//     Term 39 (AT2202-0500)/CC Outputs/Current setpoint value Ch.25 <-> Data Pointer/CurrentSetpointValues[24]
//     Term 39 (AT2202-0500)/CC Outputs/Current setpoint value Ch.26 <-> Data Pointer/CurrentSetpointValues[25]
//     Term 39 (AT2202-0500)/CC Outputs/Current setpoint value Ch.27 <-> Data Pointer/CurrentSetpointValues[26]
//     Term 39 (AT2202-0500)/CC Outputs/Current setpoint value Ch.28 <-> Data Pointer/CurrentSetpointValues[27]
//     Term 39 (AT2202-0500)/CC Outputs/Current setpoint value Ch.29 <-> Data Pointer/CurrentSetpointValues[28]
//     Term 39 (AT2202-0500)/CC Outputs/Current setpoint value Ch.3 <-> Data Pointer/CurrentSetpointValues[2]
//     Term 39 (AT2202-0500)/CC Outputs/Current setpoint value Ch.30 <-> Data Pointer/CurrentSetpointValues[29]
//     Term 39 (AT2202-0500)/CC Outputs/Current setpoint value Ch.4 <-> Data Pointer/CurrentSetpointValues[3]
//     Term 39 (AT2202-0500)/CC Outputs/Current setpoint value Ch.5 <-> Data Pointer/CurrentSetpointValues[4]
//     Term 39 (AT2202-0500)/CC Outputs/Current setpoint value Ch.6 <-> Data Pointer/CurrentSetpointValues[5]
//     Term 39 (AT2202-0500)/CC Outputs/Current setpoint value Ch.7 <-> Data Pointer/CurrentSetpointValues[6]
//     Term 39 (AT2202-0500)/CC Outputs/Current setpoint value Ch.8 <-> Data Pointer/CurrentSetpointValues[7]
//     Term 39 (AT2202-0500)/CC Outputs/Current setpoint value Ch.9 <-> Data Pointer/CurrentSetpointValues[8]
//     Term 39 (AT2202-0500)/LFB Inputs/BinaryData <-> Data Pointer/HallSensorValues
//   Device 38 <-> TcCOM Objects/XTS ProcessingUnit 1/Part 1/Module 47
//     Term 40 (AT2200-0500)/CC Inputs/Current actual value Ch.1 <-> Data Pointer/CurrentActualValues[0]
//     Term 40 (AT2200-0500)/CC Inputs/Current actual value Ch.10 <-> Data Pointer/CurrentActualValues[9]
//     Term 40 (AT2200-0500)/CC Inputs/Current actual value Ch.11 <-> Data Pointer/CurrentActualValues[10]
//     Term 40 (AT2200-0500)/CC Inputs/Current actual value Ch.12 <-> Data Pointer/CurrentActualValues[11]
//     Term 40 (AT2200-0500)/CC Inputs/Current actual value Ch.13 <-> Data Pointer/CurrentActualValues[12]
//     Term 40 (AT2200-0500)/CC Inputs/Current actual value Ch.14 <-> Data Pointer/CurrentActualValues[13]
//     Term 40 (AT2200-0500)/CC Inputs/Current actual value Ch.15 <-> Data Pointer/CurrentActualValues[14]
//     Term 40 (AT2200-0500)/CC Inputs/Current actual value Ch.16 <-> Data Pointer/CurrentActualValues[15]
//     Term 40 (AT2200-0500)/CC Inputs/Current actual value Ch.17 <-> Data Pointer/CurrentActualValues[16]
//     Term 40 (AT2200-0500)/CC Inputs/Current actual value Ch.18 <-> Data Pointer/CurrentActualValues[17]
//     Term 40 (AT2200-0500)/CC Inputs/Current actual value Ch.19 <-> Data Pointer/CurrentActualValues[18]
//     Term 40 (AT2200-0500)/CC Inputs/Current actual value Ch.2 <-> Data Pointer/CurrentActualValues[1]
//     Term 40 (AT2200-0500)/CC Inputs/Current actual value Ch.20 <-> Data Pointer/CurrentActualValues[19]
//     Term 40 (AT2200-0500)/CC Inputs/Current actual value Ch.21 <-> Data Pointer/CurrentActualValues[20]
//     Term 40 (AT2200-0500)/CC Inputs/Current actual value Ch.22 <-> Data Pointer/CurrentActualValues[21]
//     Term 40 (AT2200-0500)/CC Inputs/Current actual value Ch.23 <-> Data Pointer/CurrentActualValues[22]
//     Term 40 (AT2200-0500)/CC Inputs/Current actual value Ch.24 <-> Data Pointer/CurrentActualValues[23]
//     Term 40 (AT2200-0500)/CC Inputs/Current actual value Ch.25 <-> Data Pointer/CurrentActualValues[24]
//     Term 40 (AT2200-0500)/CC Inputs/Current actual value Ch.26 <-> Data Pointer/CurrentActualValues[25]
//     Term 40 (AT2200-0500)/CC Inputs/Current actual value Ch.27 <-> Data Pointer/CurrentActualValues[26]
//     Term 40 (AT2200-0500)/CC Inputs/Current actual value Ch.28 <-> Data Pointer/CurrentActualValues[27]
//     Term 40 (AT2200-0500)/CC Inputs/Current actual value Ch.29 <-> Data Pointer/CurrentActualValues[28]
//     Term 40 (AT2200-0500)/CC Inputs/Current actual value Ch.3 <-> Data Pointer/CurrentActualValues[2]
//     Term 40 (AT2200-0500)/CC Inputs/Current actual value Ch.30 <-> Data Pointer/CurrentActualValues[29]
//     Term 40 (AT2200-0500)/CC Inputs/Current actual value Ch.4 <-> Data Pointer/CurrentActualValues[3]
//     Term 40 (AT2200-0500)/CC Inputs/Current actual value Ch.5 <-> Data Pointer/CurrentActualValues[4]
//     Term 40 (AT2200-0500)/CC Inputs/Current actual value Ch.6 <-> Data Pointer/CurrentActualValues[5]
//     Term 40 (AT2200-0500)/CC Inputs/Current actual value Ch.7 <-> Data Pointer/CurrentActualValues[6]
//     Term 40 (AT2200-0500)/CC Inputs/Current actual value Ch.8 <-> Data Pointer/CurrentActualValues[7]
//     Term 40 (AT2200-0500)/CC Inputs/Current actual value Ch.9 <-> Data Pointer/CurrentActualValues[8]
//     Term 40 (AT2200-0500)/CC Inputs/Status <-> Data Pointer/Status
//     Term 40 (AT2200-0500)/CC Outputs/Control <-> Data Pointer/Control
//     Term 40 (AT2200-0500)/CC Outputs/Current setpoint value Ch.1 <-> Data Pointer/CurrentSetpointValues[0]
//     Term 40 (AT2200-0500)/CC Outputs/Current setpoint value Ch.10 <-> Data Pointer/CurrentSetpointValues[9]
//     Term 40 (AT2200-0500)/CC Outputs/Current setpoint value Ch.11 <-> Data Pointer/CurrentSetpointValues[10]
//     Term 40 (AT2200-0500)/CC Outputs/Current setpoint value Ch.12 <-> Data Pointer/CurrentSetpointValues[11]
//     Term 40 (AT2200-0500)/CC Outputs/Current setpoint value Ch.13 <-> Data Pointer/CurrentSetpointValues[12]
//     Term 40 (AT2200-0500)/CC Outputs/Current setpoint value Ch.14 <-> Data Pointer/CurrentSetpointValues[13]
//     Term 40 (AT2200-0500)/CC Outputs/Current setpoint value Ch.15 <-> Data Pointer/CurrentSetpointValues[14]
//     Term 40 (AT2200-0500)/CC Outputs/Current setpoint value Ch.16 <-> Data Pointer/CurrentSetpointValues[15]
//     Term 40 (AT2200-0500)/CC Outputs/Current setpoint value Ch.17 <-> Data Pointer/CurrentSetpointValues[16]
//     Term 40 (AT2200-0500)/CC Outputs/Current setpoint value Ch.18 <-> Data Pointer/CurrentSetpointValues[17]
//     Term 40 (AT2200-0500)/CC Outputs/Current setpoint value Ch.19 <-> Data Pointer/CurrentSetpointValues[18]
//     Term 40 (AT2200-0500)/CC Outputs/Current setpoint value Ch.2 <-> Data Pointer/CurrentSetpointValues[1]
//     Term 40 (AT2200-0500)/CC Outputs/Current setpoint value Ch.20 <-> Data Pointer/CurrentSetpointValues[19]
//     Term 40 (AT2200-0500)/CC Outputs/Current setpoint value Ch.21 <-> Data Pointer/CurrentSetpointValues[20]
//     Term 40 (AT2200-0500)/CC Outputs/Current setpoint value Ch.22 <-> Data Pointer/CurrentSetpointValues[21]
//     Term 40 (AT2200-0500)/CC Outputs/Current setpoint value Ch.23 <-> Data Pointer/CurrentSetpointValues[22]
//     Term 40 (AT2200-0500)/CC Outputs/Current setpoint value Ch.24 <-> Data Pointer/CurrentSetpointValues[23]
//     Term 40 (AT2200-0500)/CC Outputs/Current setpoint value Ch.25 <-> Data Pointer/CurrentSetpointValues[24]
//     Term 40 (AT2200-0500)/CC Outputs/Current setpoint value Ch.26 <-> Data Pointer/CurrentSetpointValues[25]
//     Term 40 (AT2200-0500)/CC Outputs/Current setpoint value Ch.27 <-> Data Pointer/CurrentSetpointValues[26]
//     Term 40 (AT2200-0500)/CC Outputs/Current setpoint value Ch.28 <-> Data Pointer/CurrentSetpointValues[27]
//     Term 40 (AT2200-0500)/CC Outputs/Current setpoint value Ch.29 <-> Data Pointer/CurrentSetpointValues[28]
//     Term 40 (AT2200-0500)/CC Outputs/Current setpoint value Ch.3 <-> Data Pointer/CurrentSetpointValues[2]
//     Term 40 (AT2200-0500)/CC Outputs/Current setpoint value Ch.30 <-> Data Pointer/CurrentSetpointValues[29]
//     Term 40 (AT2200-0500)/CC Outputs/Current setpoint value Ch.4 <-> Data Pointer/CurrentSetpointValues[3]
//     Term 40 (AT2200-0500)/CC Outputs/Current setpoint value Ch.5 <-> Data Pointer/CurrentSetpointValues[4]
//     Term 40 (AT2200-0500)/CC Outputs/Current setpoint value Ch.6 <-> Data Pointer/CurrentSetpointValues[5]
//     Term 40 (AT2200-0500)/CC Outputs/Current setpoint value Ch.7 <-> Data Pointer/CurrentSetpointValues[6]
//     Term 40 (AT2200-0500)/CC Outputs/Current setpoint value Ch.8 <-> Data Pointer/CurrentSetpointValues[7]
//     Term 40 (AT2200-0500)/CC Outputs/Current setpoint value Ch.9 <-> Data Pointer/CurrentSetpointValues[8]
//     Term 40 (AT2200-0500)/LFB Inputs/BinaryData <-> Data Pointer/HallSensorValues
//   Device 38 <-> TcCOM Objects/XTS ProcessingUnit 1/Part 1/Module 48
//     Term 41 (AT2200-0500)/CC Inputs/Current actual value Ch.1 <-> Data Pointer/CurrentActualValues[0]
//     Term 41 (AT2200-0500)/CC Inputs/Current actual value Ch.10 <-> Data Pointer/CurrentActualValues[9]
//     Term 41 (AT2200-0500)/CC Inputs/Current actual value Ch.11 <-> Data Pointer/CurrentActualValues[10]
//     Term 41 (AT2200-0500)/CC Inputs/Current actual value Ch.12 <-> Data Pointer/CurrentActualValues[11]
//     Term 41 (AT2200-0500)/CC Inputs/Current actual value Ch.13 <-> Data Pointer/CurrentActualValues[12]
//     Term 41 (AT2200-0500)/CC Inputs/Current actual value Ch.14 <-> Data Pointer/CurrentActualValues[13]
//     Term 41 (AT2200-0500)/CC Inputs/Current actual value Ch.15 <-> Data Pointer/CurrentActualValues[14]
//     Term 41 (AT2200-0500)/CC Inputs/Current actual value Ch.16 <-> Data Pointer/CurrentActualValues[15]
//     Term 41 (AT2200-0500)/CC Inputs/Current actual value Ch.17 <-> Data Pointer/CurrentActualValues[16]
//     Term 41 (AT2200-0500)/CC Inputs/Current actual value Ch.18 <-> Data Pointer/CurrentActualValues[17]
//     Term 41 (AT2200-0500)/CC Inputs/Current actual value Ch.19 <-> Data Pointer/CurrentActualValues[18]
//     Term 41 (AT2200-0500)/CC Inputs/Current actual value Ch.2 <-> Data Pointer/CurrentActualValues[1]
//     Term 41 (AT2200-0500)/CC Inputs/Current actual value Ch.20 <-> Data Pointer/CurrentActualValues[19]
//     Term 41 (AT2200-0500)/CC Inputs/Current actual value Ch.21 <-> Data Pointer/CurrentActualValues[20]
//     Term 41 (AT2200-0500)/CC Inputs/Current actual value Ch.22 <-> Data Pointer/CurrentActualValues[21]
//     Term 41 (AT2200-0500)/CC Inputs/Current actual value Ch.23 <-> Data Pointer/CurrentActualValues[22]
//     Term 41 (AT2200-0500)/CC Inputs/Current actual value Ch.24 <-> Data Pointer/CurrentActualValues[23]
//     Term 41 (AT2200-0500)/CC Inputs/Current actual value Ch.25 <-> Data Pointer/CurrentActualValues[24]
//     Term 41 (AT2200-0500)/CC Inputs/Current actual value Ch.26 <-> Data Pointer/CurrentActualValues[25]
//     Term 41 (AT2200-0500)/CC Inputs/Current actual value Ch.27 <-> Data Pointer/CurrentActualValues[26]
//     Term 41 (AT2200-0500)/CC Inputs/Current actual value Ch.28 <-> Data Pointer/CurrentActualValues[27]
//     Term 41 (AT2200-0500)/CC Inputs/Current actual value Ch.29 <-> Data Pointer/CurrentActualValues[28]
//     Term 41 (AT2200-0500)/CC Inputs/Current actual value Ch.3 <-> Data Pointer/CurrentActualValues[2]
//     Term 41 (AT2200-0500)/CC Inputs/Current actual value Ch.30 <-> Data Pointer/CurrentActualValues[29]
//     Term 41 (AT2200-0500)/CC Inputs/Current actual value Ch.4 <-> Data Pointer/CurrentActualValues[3]
//     Term 41 (AT2200-0500)/CC Inputs/Current actual value Ch.5 <-> Data Pointer/CurrentActualValues[4]
//     Term 41 (AT2200-0500)/CC Inputs/Current actual value Ch.6 <-> Data Pointer/CurrentActualValues[5]
//     Term 41 (AT2200-0500)/CC Inputs/Current actual value Ch.7 <-> Data Pointer/CurrentActualValues[6]
//     Term 41 (AT2200-0500)/CC Inputs/Current actual value Ch.8 <-> Data Pointer/CurrentActualValues[7]
//     Term 41 (AT2200-0500)/CC Inputs/Current actual value Ch.9 <-> Data Pointer/CurrentActualValues[8]
//     Term 41 (AT2200-0500)/CC Inputs/Status <-> Data Pointer/Status
//     Term 41 (AT2200-0500)/CC Outputs/Control <-> Data Pointer/Control
//     Term 41 (AT2200-0500)/CC Outputs/Current setpoint value Ch.1 <-> Data Pointer/CurrentSetpointValues[0]
//     Term 41 (AT2200-0500)/CC Outputs/Current setpoint value Ch.10 <-> Data Pointer/CurrentSetpointValues[9]
//     Term 41 (AT2200-0500)/CC Outputs/Current setpoint value Ch.11 <-> Data Pointer/CurrentSetpointValues[10]
//     Term 41 (AT2200-0500)/CC Outputs/Current setpoint value Ch.12 <-> Data Pointer/CurrentSetpointValues[11]
//     Term 41 (AT2200-0500)/CC Outputs/Current setpoint value Ch.13 <-> Data Pointer/CurrentSetpointValues[12]
//     Term 41 (AT2200-0500)/CC Outputs/Current setpoint value Ch.14 <-> Data Pointer/CurrentSetpointValues[13]
//     Term 41 (AT2200-0500)/CC Outputs/Current setpoint value Ch.15 <-> Data Pointer/CurrentSetpointValues[14]
//     Term 41 (AT2200-0500)/CC Outputs/Current setpoint value Ch.16 <-> Data Pointer/CurrentSetpointValues[15]
//     Term 41 (AT2200-0500)/CC Outputs/Current setpoint value Ch.17 <-> Data Pointer/CurrentSetpointValues[16]
//     Term 41 (AT2200-0500)/CC Outputs/Current setpoint value Ch.18 <-> Data Pointer/CurrentSetpointValues[17]
//     Term 41 (AT2200-0500)/CC Outputs/Current setpoint value Ch.19 <-> Data Pointer/CurrentSetpointValues[18]
//     Term 41 (AT2200-0500)/CC Outputs/Current setpoint value Ch.2 <-> Data Pointer/CurrentSetpointValues[1]
//     Term 41 (AT2200-0500)/CC Outputs/Current setpoint value Ch.20 <-> Data Pointer/CurrentSetpointValues[19]
//     Term 41 (AT2200-0500)/CC Outputs/Current setpoint value Ch.21 <-> Data Pointer/CurrentSetpointValues[20]
//     Term 41 (AT2200-0500)/CC Outputs/Current setpoint value Ch.22 <-> Data Pointer/CurrentSetpointValues[21]
//     Term 41 (AT2200-0500)/CC Outputs/Current setpoint value Ch.23 <-> Data Pointer/CurrentSetpointValues[22]
//     Term 41 (AT2200-0500)/CC Outputs/Current setpoint value Ch.24 <-> Data Pointer/CurrentSetpointValues[23]
//     Term 41 (AT2200-0500)/CC Outputs/Current setpoint value Ch.25 <-> Data Pointer/CurrentSetpointValues[24]
//     Term 41 (AT2200-0500)/CC Outputs/Current setpoint value Ch.26 <-> Data Pointer/CurrentSetpointValues[25]
//     Term 41 (AT2200-0500)/CC Outputs/Current setpoint value Ch.27 <-> Data Pointer/CurrentSetpointValues[26]
//     Term 41 (AT2200-0500)/CC Outputs/Current setpoint value Ch.28 <-> Data Pointer/CurrentSetpointValues[27]
//     Term 41 (AT2200-0500)/CC Outputs/Current setpoint value Ch.29 <-> Data Pointer/CurrentSetpointValues[28]
//     Term 41 (AT2200-0500)/CC Outputs/Current setpoint value Ch.3 <-> Data Pointer/CurrentSetpointValues[2]
//     Term 41 (AT2200-0500)/CC Outputs/Current setpoint value Ch.30 <-> Data Pointer/CurrentSetpointValues[29]
//     Term 41 (AT2200-0500)/CC Outputs/Current setpoint value Ch.4 <-> Data Pointer/CurrentSetpointValues[3]
//     Term 41 (AT2200-0500)/CC Outputs/Current setpoint value Ch.5 <-> Data Pointer/CurrentSetpointValues[4]
//     Term 41 (AT2200-0500)/CC Outputs/Current setpoint value Ch.6 <-> Data Pointer/CurrentSetpointValues[5]
//     Term 41 (AT2200-0500)/CC Outputs/Current setpoint value Ch.7 <-> Data Pointer/CurrentSetpointValues[6]
//     Term 41 (AT2200-0500)/CC Outputs/Current setpoint value Ch.8 <-> Data Pointer/CurrentSetpointValues[7]
//     Term 41 (AT2200-0500)/CC Outputs/Current setpoint value Ch.9 <-> Data Pointer/CurrentSetpointValues[8]
//     Term 41 (AT2200-0500)/LFB Inputs/BinaryData <-> Data Pointer/HallSensorValues
//   Device 39 <-> TcCOM Objects/XTS ProcessingUnit 1/Part 1/Module 49
//     Term 42 (AT2202-0500)/CC Inputs/Current actual value Ch.1 <-> Data Pointer/CurrentActualValues[0]
//     Term 42 (AT2202-0500)/CC Inputs/Current actual value Ch.10 <-> Data Pointer/CurrentActualValues[9]
//     Term 42 (AT2202-0500)/CC Inputs/Current actual value Ch.11 <-> Data Pointer/CurrentActualValues[10]
//     Term 42 (AT2202-0500)/CC Inputs/Current actual value Ch.12 <-> Data Pointer/CurrentActualValues[11]
//     Term 42 (AT2202-0500)/CC Inputs/Current actual value Ch.13 <-> Data Pointer/CurrentActualValues[12]
//     Term 42 (AT2202-0500)/CC Inputs/Current actual value Ch.14 <-> Data Pointer/CurrentActualValues[13]
//     Term 42 (AT2202-0500)/CC Inputs/Current actual value Ch.15 <-> Data Pointer/CurrentActualValues[14]
//     Term 42 (AT2202-0500)/CC Inputs/Current actual value Ch.16 <-> Data Pointer/CurrentActualValues[15]
//     Term 42 (AT2202-0500)/CC Inputs/Current actual value Ch.17 <-> Data Pointer/CurrentActualValues[16]
//     Term 42 (AT2202-0500)/CC Inputs/Current actual value Ch.18 <-> Data Pointer/CurrentActualValues[17]
//     Term 42 (AT2202-0500)/CC Inputs/Current actual value Ch.19 <-> Data Pointer/CurrentActualValues[18]
//     Term 42 (AT2202-0500)/CC Inputs/Current actual value Ch.2 <-> Data Pointer/CurrentActualValues[1]
//     Term 42 (AT2202-0500)/CC Inputs/Current actual value Ch.20 <-> Data Pointer/CurrentActualValues[19]
//     Term 42 (AT2202-0500)/CC Inputs/Current actual value Ch.21 <-> Data Pointer/CurrentActualValues[20]
//     Term 42 (AT2202-0500)/CC Inputs/Current actual value Ch.22 <-> Data Pointer/CurrentActualValues[21]
//     Term 42 (AT2202-0500)/CC Inputs/Current actual value Ch.23 <-> Data Pointer/CurrentActualValues[22]
//     Term 42 (AT2202-0500)/CC Inputs/Current actual value Ch.24 <-> Data Pointer/CurrentActualValues[23]
//     Term 42 (AT2202-0500)/CC Inputs/Current actual value Ch.25 <-> Data Pointer/CurrentActualValues[24]
//     Term 42 (AT2202-0500)/CC Inputs/Current actual value Ch.26 <-> Data Pointer/CurrentActualValues[25]
//     Term 42 (AT2202-0500)/CC Inputs/Current actual value Ch.27 <-> Data Pointer/CurrentActualValues[26]
//     Term 42 (AT2202-0500)/CC Inputs/Current actual value Ch.28 <-> Data Pointer/CurrentActualValues[27]
//     Term 42 (AT2202-0500)/CC Inputs/Current actual value Ch.29 <-> Data Pointer/CurrentActualValues[28]
//     Term 42 (AT2202-0500)/CC Inputs/Current actual value Ch.3 <-> Data Pointer/CurrentActualValues[2]
//     Term 42 (AT2202-0500)/CC Inputs/Current actual value Ch.30 <-> Data Pointer/CurrentActualValues[29]
//     Term 42 (AT2202-0500)/CC Inputs/Current actual value Ch.4 <-> Data Pointer/CurrentActualValues[3]
//     Term 42 (AT2202-0500)/CC Inputs/Current actual value Ch.5 <-> Data Pointer/CurrentActualValues[4]
//     Term 42 (AT2202-0500)/CC Inputs/Current actual value Ch.6 <-> Data Pointer/CurrentActualValues[5]
//     Term 42 (AT2202-0500)/CC Inputs/Current actual value Ch.7 <-> Data Pointer/CurrentActualValues[6]
//     Term 42 (AT2202-0500)/CC Inputs/Current actual value Ch.8 <-> Data Pointer/CurrentActualValues[7]
//     Term 42 (AT2202-0500)/CC Inputs/Current actual value Ch.9 <-> Data Pointer/CurrentActualValues[8]
//     Term 42 (AT2202-0500)/CC Inputs/Status <-> Data Pointer/Status
//     Term 42 (AT2202-0500)/CC Outputs/Control <-> Data Pointer/Control
//     Term 42 (AT2202-0500)/CC Outputs/Current setpoint value Ch.1 <-> Data Pointer/CurrentSetpointValues[0]
//     Term 42 (AT2202-0500)/CC Outputs/Current setpoint value Ch.10 <-> Data Pointer/CurrentSetpointValues[9]
//     Term 42 (AT2202-0500)/CC Outputs/Current setpoint value Ch.11 <-> Data Pointer/CurrentSetpointValues[10]
//     Term 42 (AT2202-0500)/CC Outputs/Current setpoint value Ch.12 <-> Data Pointer/CurrentSetpointValues[11]
//     Term 42 (AT2202-0500)/CC Outputs/Current setpoint value Ch.13 <-> Data Pointer/CurrentSetpointValues[12]
//     Term 42 (AT2202-0500)/CC Outputs/Current setpoint value Ch.14 <-> Data Pointer/CurrentSetpointValues[13]
//     Term 42 (AT2202-0500)/CC Outputs/Current setpoint value Ch.15 <-> Data Pointer/CurrentSetpointValues[14]
//     Term 42 (AT2202-0500)/CC Outputs/Current setpoint value Ch.16 <-> Data Pointer/CurrentSetpointValues[15]
//     Term 42 (AT2202-0500)/CC Outputs/Current setpoint value Ch.17 <-> Data Pointer/CurrentSetpointValues[16]
//     Term 42 (AT2202-0500)/CC Outputs/Current setpoint value Ch.18 <-> Data Pointer/CurrentSetpointValues[17]
//     Term 42 (AT2202-0500)/CC Outputs/Current setpoint value Ch.19 <-> Data Pointer/CurrentSetpointValues[18]
//     Term 42 (AT2202-0500)/CC Outputs/Current setpoint value Ch.2 <-> Data Pointer/CurrentSetpointValues[1]
//     Term 42 (AT2202-0500)/CC Outputs/Current setpoint value Ch.20 <-> Data Pointer/CurrentSetpointValues[19]
//     Term 42 (AT2202-0500)/CC Outputs/Current setpoint value Ch.21 <-> Data Pointer/CurrentSetpointValues[20]
//     Term 42 (AT2202-0500)/CC Outputs/Current setpoint value Ch.22 <-> Data Pointer/CurrentSetpointValues[21]
//     Term 42 (AT2202-0500)/CC Outputs/Current setpoint value Ch.23 <-> Data Pointer/CurrentSetpointValues[22]
//     Term 42 (AT2202-0500)/CC Outputs/Current setpoint value Ch.24 <-> Data Pointer/CurrentSetpointValues[23]
//     Term 42 (AT2202-0500)/CC Outputs/Current setpoint value Ch.25 <-> Data Pointer/CurrentSetpointValues[24]
//     Term 42 (AT2202-0500)/CC Outputs/Current setpoint value Ch.26 <-> Data Pointer/CurrentSetpointValues[25]
//     Term 42 (AT2202-0500)/CC Outputs/Current setpoint value Ch.27 <-> Data Pointer/CurrentSetpointValues[26]
//     Term 42 (AT2202-0500)/CC Outputs/Current setpoint value Ch.28 <-> Data Pointer/CurrentSetpointValues[27]
//     Term 42 (AT2202-0500)/CC Outputs/Current setpoint value Ch.29 <-> Data Pointer/CurrentSetpointValues[28]
//     Term 42 (AT2202-0500)/CC Outputs/Current setpoint value Ch.3 <-> Data Pointer/CurrentSetpointValues[2]
//     Term 42 (AT2202-0500)/CC Outputs/Current setpoint value Ch.30 <-> Data Pointer/CurrentSetpointValues[29]
//     Term 42 (AT2202-0500)/CC Outputs/Current setpoint value Ch.4 <-> Data Pointer/CurrentSetpointValues[3]
//     Term 42 (AT2202-0500)/CC Outputs/Current setpoint value Ch.5 <-> Data Pointer/CurrentSetpointValues[4]
//     Term 42 (AT2202-0500)/CC Outputs/Current setpoint value Ch.6 <-> Data Pointer/CurrentSetpointValues[5]
//     Term 42 (AT2202-0500)/CC Outputs/Current setpoint value Ch.7 <-> Data Pointer/CurrentSetpointValues[6]
//     Term 42 (AT2202-0500)/CC Outputs/Current setpoint value Ch.8 <-> Data Pointer/CurrentSetpointValues[7]
//     Term 42 (AT2202-0500)/CC Outputs/Current setpoint value Ch.9 <-> Data Pointer/CurrentSetpointValues[8]
//     Term 42 (AT2202-0500)/LFB Inputs/BinaryData <-> Data Pointer/HallSensorValues
//   Device 39 <-> TcCOM Objects/XTS ProcessingUnit 1/Part 1/Module 50
//     Term 43 (AT2200-0500)/CC Inputs/Current actual value Ch.1 <-> Data Pointer/CurrentActualValues[0]
//     Term 43 (AT2200-0500)/CC Inputs/Current actual value Ch.10 <-> Data Pointer/CurrentActualValues[9]
//     Term 43 (AT2200-0500)/CC Inputs/Current actual value Ch.11 <-> Data Pointer/CurrentActualValues[10]
//     Term 43 (AT2200-0500)/CC Inputs/Current actual value Ch.12 <-> Data Pointer/CurrentActualValues[11]
//     Term 43 (AT2200-0500)/CC Inputs/Current actual value Ch.13 <-> Data Pointer/CurrentActualValues[12]
//     Term 43 (AT2200-0500)/CC Inputs/Current actual value Ch.14 <-> Data Pointer/CurrentActualValues[13]
//     Term 43 (AT2200-0500)/CC Inputs/Current actual value Ch.15 <-> Data Pointer/CurrentActualValues[14]
//     Term 43 (AT2200-0500)/CC Inputs/Current actual value Ch.16 <-> Data Pointer/CurrentActualValues[15]
//     Term 43 (AT2200-0500)/CC Inputs/Current actual value Ch.17 <-> Data Pointer/CurrentActualValues[16]
//     Term 43 (AT2200-0500)/CC Inputs/Current actual value Ch.18 <-> Data Pointer/CurrentActualValues[17]
//     Term 43 (AT2200-0500)/CC Inputs/Current actual value Ch.19 <-> Data Pointer/CurrentActualValues[18]
//     Term 43 (AT2200-0500)/CC Inputs/Current actual value Ch.2 <-> Data Pointer/CurrentActualValues[1]
//     Term 43 (AT2200-0500)/CC Inputs/Current actual value Ch.20 <-> Data Pointer/CurrentActualValues[19]
//     Term 43 (AT2200-0500)/CC Inputs/Current actual value Ch.21 <-> Data Pointer/CurrentActualValues[20]
//     Term 43 (AT2200-0500)/CC Inputs/Current actual value Ch.22 <-> Data Pointer/CurrentActualValues[21]
//     Term 43 (AT2200-0500)/CC Inputs/Current actual value Ch.23 <-> Data Pointer/CurrentActualValues[22]
//     Term 43 (AT2200-0500)/CC Inputs/Current actual value Ch.24 <-> Data Pointer/CurrentActualValues[23]
//     Term 43 (AT2200-0500)/CC Inputs/Current actual value Ch.25 <-> Data Pointer/CurrentActualValues[24]
//     Term 43 (AT2200-0500)/CC Inputs/Current actual value Ch.26 <-> Data Pointer/CurrentActualValues[25]
//     Term 43 (AT2200-0500)/CC Inputs/Current actual value Ch.27 <-> Data Pointer/CurrentActualValues[26]
//     Term 43 (AT2200-0500)/CC Inputs/Current actual value Ch.28 <-> Data Pointer/CurrentActualValues[27]
//     Term 43 (AT2200-0500)/CC Inputs/Current actual value Ch.29 <-> Data Pointer/CurrentActualValues[28]
//     Term 43 (AT2200-0500)/CC Inputs/Current actual value Ch.3 <-> Data Pointer/CurrentActualValues[2]
//     Term 43 (AT2200-0500)/CC Inputs/Current actual value Ch.30 <-> Data Pointer/CurrentActualValues[29]
//     Term 43 (AT2200-0500)/CC Inputs/Current actual value Ch.4 <-> Data Pointer/CurrentActualValues[3]
//     Term 43 (AT2200-0500)/CC Inputs/Current actual value Ch.5 <-> Data Pointer/CurrentActualValues[4]
//     Term 43 (AT2200-0500)/CC Inputs/Current actual value Ch.6 <-> Data Pointer/CurrentActualValues[5]
//     Term 43 (AT2200-0500)/CC Inputs/Current actual value Ch.7 <-> Data Pointer/CurrentActualValues[6]
//     Term 43 (AT2200-0500)/CC Inputs/Current actual value Ch.8 <-> Data Pointer/CurrentActualValues[7]
//     Term 43 (AT2200-0500)/CC Inputs/Current actual value Ch.9 <-> Data Pointer/CurrentActualValues[8]
//     Term 43 (AT2200-0500)/CC Inputs/Status <-> Data Pointer/Status
//     Term 43 (AT2200-0500)/CC Outputs/Control <-> Data Pointer/Control
//     Term 43 (AT2200-0500)/CC Outputs/Current setpoint value Ch.1 <-> Data Pointer/CurrentSetpointValues[0]
//     Term 43 (AT2200-0500)/CC Outputs/Current setpoint value Ch.10 <-> Data Pointer/CurrentSetpointValues[9]
//     Term 43 (AT2200-0500)/CC Outputs/Current setpoint value Ch.11 <-> Data Pointer/CurrentSetpointValues[10]
//     Term 43 (AT2200-0500)/CC Outputs/Current setpoint value Ch.12 <-> Data Pointer/CurrentSetpointValues[11]
//     Term 43 (AT2200-0500)/CC Outputs/Current setpoint value Ch.13 <-> Data Pointer/CurrentSetpointValues[12]
//     Term 43 (AT2200-0500)/CC Outputs/Current setpoint value Ch.14 <-> Data Pointer/CurrentSetpointValues[13]
//     Term 43 (AT2200-0500)/CC Outputs/Current setpoint value Ch.15 <-> Data Pointer/CurrentSetpointValues[14]
//     Term 43 (AT2200-0500)/CC Outputs/Current setpoint value Ch.16 <-> Data Pointer/CurrentSetpointValues[15]
//     Term 43 (AT2200-0500)/CC Outputs/Current setpoint value Ch.17 <-> Data Pointer/CurrentSetpointValues[16]
//     Term 43 (AT2200-0500)/CC Outputs/Current setpoint value Ch.18 <-> Data Pointer/CurrentSetpointValues[17]
//     Term 43 (AT2200-0500)/CC Outputs/Current setpoint value Ch.19 <-> Data Pointer/CurrentSetpointValues[18]
//     Term 43 (AT2200-0500)/CC Outputs/Current setpoint value Ch.2 <-> Data Pointer/CurrentSetpointValues[1]
//     Term 43 (AT2200-0500)/CC Outputs/Current setpoint value Ch.20 <-> Data Pointer/CurrentSetpointValues[19]
//     Term 43 (AT2200-0500)/CC Outputs/Current setpoint value Ch.21 <-> Data Pointer/CurrentSetpointValues[20]
//     Term 43 (AT2200-0500)/CC Outputs/Current setpoint value Ch.22 <-> Data Pointer/CurrentSetpointValues[21]
//     Term 43 (AT2200-0500)/CC Outputs/Current setpoint value Ch.23 <-> Data Pointer/CurrentSetpointValues[22]
//     Term 43 (AT2200-0500)/CC Outputs/Current setpoint value Ch.24 <-> Data Pointer/CurrentSetpointValues[23]
//     Term 43 (AT2200-0500)/CC Outputs/Current setpoint value Ch.25 <-> Data Pointer/CurrentSetpointValues[24]
//     Term 43 (AT2200-0500)/CC Outputs/Current setpoint value Ch.26 <-> Data Pointer/CurrentSetpointValues[25]
//     Term 43 (AT2200-0500)/CC Outputs/Current setpoint value Ch.27 <-> Data Pointer/CurrentSetpointValues[26]
//     Term 43 (AT2200-0500)/CC Outputs/Current setpoint value Ch.28 <-> Data Pointer/CurrentSetpointValues[27]
//     Term 43 (AT2200-0500)/CC Outputs/Current setpoint value Ch.29 <-> Data Pointer/CurrentSetpointValues[28]
//     Term 43 (AT2200-0500)/CC Outputs/Current setpoint value Ch.3 <-> Data Pointer/CurrentSetpointValues[2]
//     Term 43 (AT2200-0500)/CC Outputs/Current setpoint value Ch.30 <-> Data Pointer/CurrentSetpointValues[29]
//     Term 43 (AT2200-0500)/CC Outputs/Current setpoint value Ch.4 <-> Data Pointer/CurrentSetpointValues[3]
//     Term 43 (AT2200-0500)/CC Outputs/Current setpoint value Ch.5 <-> Data Pointer/CurrentSetpointValues[4]
//     Term 43 (AT2200-0500)/CC Outputs/Current setpoint value Ch.6 <-> Data Pointer/CurrentSetpointValues[5]
//     Term 43 (AT2200-0500)/CC Outputs/Current setpoint value Ch.7 <-> Data Pointer/CurrentSetpointValues[6]
//     Term 43 (AT2200-0500)/CC Outputs/Current setpoint value Ch.8 <-> Data Pointer/CurrentSetpointValues[7]
//     Term 43 (AT2200-0500)/CC Outputs/Current setpoint value Ch.9 <-> Data Pointer/CurrentSetpointValues[8]
//     Term 43 (AT2200-0500)/LFB Inputs/BinaryData <-> Data Pointer/HallSensorValues
//   Device 39 <-> TcCOM Objects/XTS ProcessingUnit 1/Part 1/Module 51
//     Term 44 (AT2200-0500)/CC Inputs/Current actual value Ch.1 <-> Data Pointer/CurrentActualValues[0]
//     Term 44 (AT2200-0500)/CC Inputs/Current actual value Ch.10 <-> Data Pointer/CurrentActualValues[9]
//     Term 44 (AT2200-0500)/CC Inputs/Current actual value Ch.11 <-> Data Pointer/CurrentActualValues[10]
//     Term 44 (AT2200-0500)/CC Inputs/Current actual value Ch.12 <-> Data Pointer/CurrentActualValues[11]
//     Term 44 (AT2200-0500)/CC Inputs/Current actual value Ch.13 <-> Data Pointer/CurrentActualValues[12]
//     Term 44 (AT2200-0500)/CC Inputs/Current actual value Ch.14 <-> Data Pointer/CurrentActualValues[13]
//     Term 44 (AT2200-0500)/CC Inputs/Current actual value Ch.15 <-> Data Pointer/CurrentActualValues[14]
//     Term 44 (AT2200-0500)/CC Inputs/Current actual value Ch.16 <-> Data Pointer/CurrentActualValues[15]
//     Term 44 (AT2200-0500)/CC Inputs/Current actual value Ch.17 <-> Data Pointer/CurrentActualValues[16]
//     Term 44 (AT2200-0500)/CC Inputs/Current actual value Ch.18 <-> Data Pointer/CurrentActualValues[17]
//     Term 44 (AT2200-0500)/CC Inputs/Current actual value Ch.19 <-> Data Pointer/CurrentActualValues[18]
//     Term 44 (AT2200-0500)/CC Inputs/Current actual value Ch.2 <-> Data Pointer/CurrentActualValues[1]
//     Term 44 (AT2200-0500)/CC Inputs/Current actual value Ch.20 <-> Data Pointer/CurrentActualValues[19]
//     Term 44 (AT2200-0500)/CC Inputs/Current actual value Ch.21 <-> Data Pointer/CurrentActualValues[20]
//     Term 44 (AT2200-0500)/CC Inputs/Current actual value Ch.22 <-> Data Pointer/CurrentActualValues[21]
//     Term 44 (AT2200-0500)/CC Inputs/Current actual value Ch.23 <-> Data Pointer/CurrentActualValues[22]
//     Term 44 (AT2200-0500)/CC Inputs/Current actual value Ch.24 <-> Data Pointer/CurrentActualValues[23]
//     Term 44 (AT2200-0500)/CC Inputs/Current actual value Ch.25 <-> Data Pointer/CurrentActualValues[24]
//     Term 44 (AT2200-0500)/CC Inputs/Current actual value Ch.26 <-> Data Pointer/CurrentActualValues[25]
//     Term 44 (AT2200-0500)/CC Inputs/Current actual value Ch.27 <-> Data Pointer/CurrentActualValues[26]
//     Term 44 (AT2200-0500)/CC Inputs/Current actual value Ch.28 <-> Data Pointer/CurrentActualValues[27]
//     Term 44 (AT2200-0500)/CC Inputs/Current actual value Ch.29 <-> Data Pointer/CurrentActualValues[28]
//     Term 44 (AT2200-0500)/CC Inputs/Current actual value Ch.3 <-> Data Pointer/CurrentActualValues[2]
//     Term 44 (AT2200-0500)/CC Inputs/Current actual value Ch.30 <-> Data Pointer/CurrentActualValues[29]
//     Term 44 (AT2200-0500)/CC Inputs/Current actual value Ch.4 <-> Data Pointer/CurrentActualValues[3]
//     Term 44 (AT2200-0500)/CC Inputs/Current actual value Ch.5 <-> Data Pointer/CurrentActualValues[4]
//     Term 44 (AT2200-0500)/CC Inputs/Current actual value Ch.6 <-> Data Pointer/CurrentActualValues[5]
//     Term 44 (AT2200-0500)/CC Inputs/Current actual value Ch.7 <-> Data Pointer/CurrentActualValues[6]
//     Term 44 (AT2200-0500)/CC Inputs/Current actual value Ch.8 <-> Data Pointer/CurrentActualValues[7]
//     Term 44 (AT2200-0500)/CC Inputs/Current actual value Ch.9 <-> Data Pointer/CurrentActualValues[8]
//     Term 44 (AT2200-0500)/CC Inputs/Status <-> Data Pointer/Status
//     Term 44 (AT2200-0500)/CC Outputs/Control <-> Data Pointer/Control
//     Term 44 (AT2200-0500)/CC Outputs/Current setpoint value Ch.1 <-> Data Pointer/CurrentSetpointValues[0]
//     Term 44 (AT2200-0500)/CC Outputs/Current setpoint value Ch.10 <-> Data Pointer/CurrentSetpointValues[9]
//     Term 44 (AT2200-0500)/CC Outputs/Current setpoint value Ch.11 <-> Data Pointer/CurrentSetpointValues[10]
//     Term 44 (AT2200-0500)/CC Outputs/Current setpoint value Ch.12 <-> Data Pointer/CurrentSetpointValues[11]
//     Term 44 (AT2200-0500)/CC Outputs/Current setpoint value Ch.13 <-> Data Pointer/CurrentSetpointValues[12]
//     Term 44 (AT2200-0500)/CC Outputs/Current setpoint value Ch.14 <-> Data Pointer/CurrentSetpointValues[13]
//     Term 44 (AT2200-0500)/CC Outputs/Current setpoint value Ch.15 <-> Data Pointer/CurrentSetpointValues[14]
//     Term 44 (AT2200-0500)/CC Outputs/Current setpoint value Ch.16 <-> Data Pointer/CurrentSetpointValues[15]
//     Term 44 (AT2200-0500)/CC Outputs/Current setpoint value Ch.17 <-> Data Pointer/CurrentSetpointValues[16]
//     Term 44 (AT2200-0500)/CC Outputs/Current setpoint value Ch.18 <-> Data Pointer/CurrentSetpointValues[17]
//     Term 44 (AT2200-0500)/CC Outputs/Current setpoint value Ch.19 <-> Data Pointer/CurrentSetpointValues[18]
//     Term 44 (AT2200-0500)/CC Outputs/Current setpoint value Ch.2 <-> Data Pointer/CurrentSetpointValues[1]
//     Term 44 (AT2200-0500)/CC Outputs/Current setpoint value Ch.20 <-> Data Pointer/CurrentSetpointValues[19]
//     Term 44 (AT2200-0500)/CC Outputs/Current setpoint value Ch.21 <-> Data Pointer/CurrentSetpointValues[20]
//     Term 44 (AT2200-0500)/CC Outputs/Current setpoint value Ch.22 <-> Data Pointer/CurrentSetpointValues[21]
//     Term 44 (AT2200-0500)/CC Outputs/Current setpoint value Ch.23 <-> Data Pointer/CurrentSetpointValues[22]
//     Term 44 (AT2200-0500)/CC Outputs/Current setpoint value Ch.24 <-> Data Pointer/CurrentSetpointValues[23]
//     Term 44 (AT2200-0500)/CC Outputs/Current setpoint value Ch.25 <-> Data Pointer/CurrentSetpointValues[24]
//     Term 44 (AT2200-0500)/CC Outputs/Current setpoint value Ch.26 <-> Data Pointer/CurrentSetpointValues[25]
//     Term 44 (AT2200-0500)/CC Outputs/Current setpoint value Ch.27 <-> Data Pointer/CurrentSetpointValues[26]
//     Term 44 (AT2200-0500)/CC Outputs/Current setpoint value Ch.28 <-> Data Pointer/CurrentSetpointValues[27]
//     Term 44 (AT2200-0500)/CC Outputs/Current setpoint value Ch.29 <-> Data Pointer/CurrentSetpointValues[28]
//     Term 44 (AT2200-0500)/CC Outputs/Current setpoint value Ch.3 <-> Data Pointer/CurrentSetpointValues[2]
//     Term 44 (AT2200-0500)/CC Outputs/Current setpoint value Ch.30 <-> Data Pointer/CurrentSetpointValues[29]
//     Term 44 (AT2200-0500)/CC Outputs/Current setpoint value Ch.4 <-> Data Pointer/CurrentSetpointValues[3]
//     Term 44 (AT2200-0500)/CC Outputs/Current setpoint value Ch.5 <-> Data Pointer/CurrentSetpointValues[4]
//     Term 44 (AT2200-0500)/CC Outputs/Current setpoint value Ch.6 <-> Data Pointer/CurrentSetpointValues[5]
//     Term 44 (AT2200-0500)/CC Outputs/Current setpoint value Ch.7 <-> Data Pointer/CurrentSetpointValues[6]
//     Term 44 (AT2200-0500)/CC Outputs/Current setpoint value Ch.8 <-> Data Pointer/CurrentSetpointValues[7]
//     Term 44 (AT2200-0500)/CC Outputs/Current setpoint value Ch.9 <-> Data Pointer/CurrentSetpointValues[8]
//     Term 44 (AT2200-0500)/LFB Inputs/BinaryData <-> Data Pointer/HallSensorValues
//   Device 40 <-> TcCOM Objects/XTS ProcessingUnit 1/Part 1/Module 52
//     Term 45 (AT2202-0500)/CC Inputs/Current actual value Ch.1 <-> Data Pointer/CurrentActualValues[0]
//     Term 45 (AT2202-0500)/CC Inputs/Current actual value Ch.10 <-> Data Pointer/CurrentActualValues[9]
//     Term 45 (AT2202-0500)/CC Inputs/Current actual value Ch.11 <-> Data Pointer/CurrentActualValues[10]
//     Term 45 (AT2202-0500)/CC Inputs/Current actual value Ch.12 <-> Data Pointer/CurrentActualValues[11]
//     Term 45 (AT2202-0500)/CC Inputs/Current actual value Ch.13 <-> Data Pointer/CurrentActualValues[12]
//     Term 45 (AT2202-0500)/CC Inputs/Current actual value Ch.14 <-> Data Pointer/CurrentActualValues[13]
//     Term 45 (AT2202-0500)/CC Inputs/Current actual value Ch.15 <-> Data Pointer/CurrentActualValues[14]
//     Term 45 (AT2202-0500)/CC Inputs/Current actual value Ch.16 <-> Data Pointer/CurrentActualValues[15]
//     Term 45 (AT2202-0500)/CC Inputs/Current actual value Ch.17 <-> Data Pointer/CurrentActualValues[16]
//     Term 45 (AT2202-0500)/CC Inputs/Current actual value Ch.18 <-> Data Pointer/CurrentActualValues[17]
//     Term 45 (AT2202-0500)/CC Inputs/Current actual value Ch.19 <-> Data Pointer/CurrentActualValues[18]
//     Term 45 (AT2202-0500)/CC Inputs/Current actual value Ch.2 <-> Data Pointer/CurrentActualValues[1]
//     Term 45 (AT2202-0500)/CC Inputs/Current actual value Ch.20 <-> Data Pointer/CurrentActualValues[19]
//     Term 45 (AT2202-0500)/CC Inputs/Current actual value Ch.21 <-> Data Pointer/CurrentActualValues[20]
//     Term 45 (AT2202-0500)/CC Inputs/Current actual value Ch.22 <-> Data Pointer/CurrentActualValues[21]
//     Term 45 (AT2202-0500)/CC Inputs/Current actual value Ch.23 <-> Data Pointer/CurrentActualValues[22]
//     Term 45 (AT2202-0500)/CC Inputs/Current actual value Ch.24 <-> Data Pointer/CurrentActualValues[23]
//     Term 45 (AT2202-0500)/CC Inputs/Current actual value Ch.25 <-> Data Pointer/CurrentActualValues[24]
//     Term 45 (AT2202-0500)/CC Inputs/Current actual value Ch.26 <-> Data Pointer/CurrentActualValues[25]
//     Term 45 (AT2202-0500)/CC Inputs/Current actual value Ch.27 <-> Data Pointer/CurrentActualValues[26]
//     Term 45 (AT2202-0500)/CC Inputs/Current actual value Ch.28 <-> Data Pointer/CurrentActualValues[27]
//     Term 45 (AT2202-0500)/CC Inputs/Current actual value Ch.29 <-> Data Pointer/CurrentActualValues[28]
//     Term 45 (AT2202-0500)/CC Inputs/Current actual value Ch.3 <-> Data Pointer/CurrentActualValues[2]
//     Term 45 (AT2202-0500)/CC Inputs/Current actual value Ch.30 <-> Data Pointer/CurrentActualValues[29]
//     Term 45 (AT2202-0500)/CC Inputs/Current actual value Ch.4 <-> Data Pointer/CurrentActualValues[3]
//     Term 45 (AT2202-0500)/CC Inputs/Current actual value Ch.5 <-> Data Pointer/CurrentActualValues[4]
//     Term 45 (AT2202-0500)/CC Inputs/Current actual value Ch.6 <-> Data Pointer/CurrentActualValues[5]
//     Term 45 (AT2202-0500)/CC Inputs/Current actual value Ch.7 <-> Data Pointer/CurrentActualValues[6]
//     Term 45 (AT2202-0500)/CC Inputs/Current actual value Ch.8 <-> Data Pointer/CurrentActualValues[7]
//     Term 45 (AT2202-0500)/CC Inputs/Current actual value Ch.9 <-> Data Pointer/CurrentActualValues[8]
//     Term 45 (AT2202-0500)/CC Inputs/Status <-> Data Pointer/Status
//     Term 45 (AT2202-0500)/CC Outputs/Control <-> Data Pointer/Control
//     Term 45 (AT2202-0500)/CC Outputs/Current setpoint value Ch.1 <-> Data Pointer/CurrentSetpointValues[0]
//     Term 45 (AT2202-0500)/CC Outputs/Current setpoint value Ch.10 <-> Data Pointer/CurrentSetpointValues[9]
//     Term 45 (AT2202-0500)/CC Outputs/Current setpoint value Ch.11 <-> Data Pointer/CurrentSetpointValues[10]
//     Term 45 (AT2202-0500)/CC Outputs/Current setpoint value Ch.12 <-> Data Pointer/CurrentSetpointValues[11]
//     Term 45 (AT2202-0500)/CC Outputs/Current setpoint value Ch.13 <-> Data Pointer/CurrentSetpointValues[12]
//     Term 45 (AT2202-0500)/CC Outputs/Current setpoint value Ch.14 <-> Data Pointer/CurrentSetpointValues[13]
//     Term 45 (AT2202-0500)/CC Outputs/Current setpoint value Ch.15 <-> Data Pointer/CurrentSetpointValues[14]
//     Term 45 (AT2202-0500)/CC Outputs/Current setpoint value Ch.16 <-> Data Pointer/CurrentSetpointValues[15]
//     Term 45 (AT2202-0500)/CC Outputs/Current setpoint value Ch.17 <-> Data Pointer/CurrentSetpointValues[16]
//     Term 45 (AT2202-0500)/CC Outputs/Current setpoint value Ch.18 <-> Data Pointer/CurrentSetpointValues[17]
//     Term 45 (AT2202-0500)/CC Outputs/Current setpoint value Ch.19 <-> Data Pointer/CurrentSetpointValues[18]
//     Term 45 (AT2202-0500)/CC Outputs/Current setpoint value Ch.2 <-> Data Pointer/CurrentSetpointValues[1]
//     Term 45 (AT2202-0500)/CC Outputs/Current setpoint value Ch.20 <-> Data Pointer/CurrentSetpointValues[19]
//     Term 45 (AT2202-0500)/CC Outputs/Current setpoint value Ch.21 <-> Data Pointer/CurrentSetpointValues[20]
//     Term 45 (AT2202-0500)/CC Outputs/Current setpoint value Ch.22 <-> Data Pointer/CurrentSetpointValues[21]
//     Term 45 (AT2202-0500)/CC Outputs/Current setpoint value Ch.23 <-> Data Pointer/CurrentSetpointValues[22]
//     Term 45 (AT2202-0500)/CC Outputs/Current setpoint value Ch.24 <-> Data Pointer/CurrentSetpointValues[23]
//     Term 45 (AT2202-0500)/CC Outputs/Current setpoint value Ch.25 <-> Data Pointer/CurrentSetpointValues[24]
//     Term 45 (AT2202-0500)/CC Outputs/Current setpoint value Ch.26 <-> Data Pointer/CurrentSetpointValues[25]
//     Term 45 (AT2202-0500)/CC Outputs/Current setpoint value Ch.27 <-> Data Pointer/CurrentSetpointValues[26]
//     Term 45 (AT2202-0500)/CC Outputs/Current setpoint value Ch.28 <-> Data Pointer/CurrentSetpointValues[27]
//     Term 45 (AT2202-0500)/CC Outputs/Current setpoint value Ch.29 <-> Data Pointer/CurrentSetpointValues[28]
//     Term 45 (AT2202-0500)/CC Outputs/Current setpoint value Ch.3 <-> Data Pointer/CurrentSetpointValues[2]
//     Term 45 (AT2202-0500)/CC Outputs/Current setpoint value Ch.30 <-> Data Pointer/CurrentSetpointValues[29]
//     Term 45 (AT2202-0500)/CC Outputs/Current setpoint value Ch.4 <-> Data Pointer/CurrentSetpointValues[3]
//     Term 45 (AT2202-0500)/CC Outputs/Current setpoint value Ch.5 <-> Data Pointer/CurrentSetpointValues[4]
//     Term 45 (AT2202-0500)/CC Outputs/Current setpoint value Ch.6 <-> Data Pointer/CurrentSetpointValues[5]
//     Term 45 (AT2202-0500)/CC Outputs/Current setpoint value Ch.7 <-> Data Pointer/CurrentSetpointValues[6]
//     Term 45 (AT2202-0500)/CC Outputs/Current setpoint value Ch.8 <-> Data Pointer/CurrentSetpointValues[7]
//     Term 45 (AT2202-0500)/CC Outputs/Current setpoint value Ch.9 <-> Data Pointer/CurrentSetpointValues[8]
//     Term 45 (AT2202-0500)/LFB Inputs/BinaryData <-> Data Pointer/HallSensorValues
//   Device 40 <-> TcCOM Objects/XTS ProcessingUnit 1/Part 1/Module 53
//     Term 46 (AT2200-0500)/CC Inputs/Current actual value Ch.1 <-> Data Pointer/CurrentActualValues[0]
//     Term 46 (AT2200-0500)/CC Inputs/Current actual value Ch.10 <-> Data Pointer/CurrentActualValues[9]
//     Term 46 (AT2200-0500)/CC Inputs/Current actual value Ch.11 <-> Data Pointer/CurrentActualValues[10]
//     Term 46 (AT2200-0500)/CC Inputs/Current actual value Ch.12 <-> Data Pointer/CurrentActualValues[11]
//     Term 46 (AT2200-0500)/CC Inputs/Current actual value Ch.13 <-> Data Pointer/CurrentActualValues[12]
//     Term 46 (AT2200-0500)/CC Inputs/Current actual value Ch.14 <-> Data Pointer/CurrentActualValues[13]
//     Term 46 (AT2200-0500)/CC Inputs/Current actual value Ch.15 <-> Data Pointer/CurrentActualValues[14]
//     Term 46 (AT2200-0500)/CC Inputs/Current actual value Ch.16 <-> Data Pointer/CurrentActualValues[15]
//     Term 46 (AT2200-0500)/CC Inputs/Current actual value Ch.17 <-> Data Pointer/CurrentActualValues[16]
//     Term 46 (AT2200-0500)/CC Inputs/Current actual value Ch.18 <-> Data Pointer/CurrentActualValues[17]
//     Term 46 (AT2200-0500)/CC Inputs/Current actual value Ch.19 <-> Data Pointer/CurrentActualValues[18]
//     Term 46 (AT2200-0500)/CC Inputs/Current actual value Ch.2 <-> Data Pointer/CurrentActualValues[1]
//     Term 46 (AT2200-0500)/CC Inputs/Current actual value Ch.20 <-> Data Pointer/CurrentActualValues[19]
//     Term 46 (AT2200-0500)/CC Inputs/Current actual value Ch.21 <-> Data Pointer/CurrentActualValues[20]
//     Term 46 (AT2200-0500)/CC Inputs/Current actual value Ch.22 <-> Data Pointer/CurrentActualValues[21]
//     Term 46 (AT2200-0500)/CC Inputs/Current actual value Ch.23 <-> Data Pointer/CurrentActualValues[22]
//     Term 46 (AT2200-0500)/CC Inputs/Current actual value Ch.24 <-> Data Pointer/CurrentActualValues[23]
//     Term 46 (AT2200-0500)/CC Inputs/Current actual value Ch.25 <-> Data Pointer/CurrentActualValues[24]
//     Term 46 (AT2200-0500)/CC Inputs/Current actual value Ch.26 <-> Data Pointer/CurrentActualValues[25]
//     Term 46 (AT2200-0500)/CC Inputs/Current actual value Ch.27 <-> Data Pointer/CurrentActualValues[26]
//     Term 46 (AT2200-0500)/CC Inputs/Current actual value Ch.28 <-> Data Pointer/CurrentActualValues[27]
//     Term 46 (AT2200-0500)/CC Inputs/Current actual value Ch.29 <-> Data Pointer/CurrentActualValues[28]
//     Term 46 (AT2200-0500)/CC Inputs/Current actual value Ch.3 <-> Data Pointer/CurrentActualValues[2]
//     Term 46 (AT2200-0500)/CC Inputs/Current actual value Ch.30 <-> Data Pointer/CurrentActualValues[29]
//     Term 46 (AT2200-0500)/CC Inputs/Current actual value Ch.4 <-> Data Pointer/CurrentActualValues[3]
//     Term 46 (AT2200-0500)/CC Inputs/Current actual value Ch.5 <-> Data Pointer/CurrentActualValues[4]
//     Term 46 (AT2200-0500)/CC Inputs/Current actual value Ch.6 <-> Data Pointer/CurrentActualValues[5]
//     Term 46 (AT2200-0500)/CC Inputs/Current actual value Ch.7 <-> Data Pointer/CurrentActualValues[6]
//     Term 46 (AT2200-0500)/CC Inputs/Current actual value Ch.8 <-> Data Pointer/CurrentActualValues[7]
//     Term 46 (AT2200-0500)/CC Inputs/Current actual value Ch.9 <-> Data Pointer/CurrentActualValues[8]
//     Term 46 (AT2200-0500)/CC Inputs/Status <-> Data Pointer/Status
//     Term 46 (AT2200-0500)/CC Outputs/Control <-> Data Pointer/Control
//     Term 46 (AT2200-0500)/CC Outputs/Current setpoint value Ch.1 <-> Data Pointer/CurrentSetpointValues[0]
//     Term 46 (AT2200-0500)/CC Outputs/Current setpoint value Ch.10 <-> Data Pointer/CurrentSetpointValues[9]
//     Term 46 (AT2200-0500)/CC Outputs/Current setpoint value Ch.11 <-> Data Pointer/CurrentSetpointValues[10]
//     Term 46 (AT2200-0500)/CC Outputs/Current setpoint value Ch.12 <-> Data Pointer/CurrentSetpointValues[11]
//     Term 46 (AT2200-0500)/CC Outputs/Current setpoint value Ch.13 <-> Data Pointer/CurrentSetpointValues[12]
//     Term 46 (AT2200-0500)/CC Outputs/Current setpoint value Ch.14 <-> Data Pointer/CurrentSetpointValues[13]
//     Term 46 (AT2200-0500)/CC Outputs/Current setpoint value Ch.15 <-> Data Pointer/CurrentSetpointValues[14]
//     Term 46 (AT2200-0500)/CC Outputs/Current setpoint value Ch.16 <-> Data Pointer/CurrentSetpointValues[15]
//     Term 46 (AT2200-0500)/CC Outputs/Current setpoint value Ch.17 <-> Data Pointer/CurrentSetpointValues[16]
//     Term 46 (AT2200-0500)/CC Outputs/Current setpoint value Ch.18 <-> Data Pointer/CurrentSetpointValues[17]
//     Term 46 (AT2200-0500)/CC Outputs/Current setpoint value Ch.19 <-> Data Pointer/CurrentSetpointValues[18]
//     Term 46 (AT2200-0500)/CC Outputs/Current setpoint value Ch.2 <-> Data Pointer/CurrentSetpointValues[1]
//     Term 46 (AT2200-0500)/CC Outputs/Current setpoint value Ch.20 <-> Data Pointer/CurrentSetpointValues[19]
//     Term 46 (AT2200-0500)/CC Outputs/Current setpoint value Ch.21 <-> Data Pointer/CurrentSetpointValues[20]
//     Term 46 (AT2200-0500)/CC Outputs/Current setpoint value Ch.22 <-> Data Pointer/CurrentSetpointValues[21]
//     Term 46 (AT2200-0500)/CC Outputs/Current setpoint value Ch.23 <-> Data Pointer/CurrentSetpointValues[22]
//     Term 46 (AT2200-0500)/CC Outputs/Current setpoint value Ch.24 <-> Data Pointer/CurrentSetpointValues[23]
//     Term 46 (AT2200-0500)/CC Outputs/Current setpoint value Ch.25 <-> Data Pointer/CurrentSetpointValues[24]
//     Term 46 (AT2200-0500)/CC Outputs/Current setpoint value Ch.26 <-> Data Pointer/CurrentSetpointValues[25]
//     Term 46 (AT2200-0500)/CC Outputs/Current setpoint value Ch.27 <-> Data Pointer/CurrentSetpointValues[26]
//     Term 46 (AT2200-0500)/CC Outputs/Current setpoint value Ch.28 <-> Data Pointer/CurrentSetpointValues[27]
//     Term 46 (AT2200-0500)/CC Outputs/Current setpoint value Ch.29 <-> Data Pointer/CurrentSetpointValues[28]
//     Term 46 (AT2200-0500)/CC Outputs/Current setpoint value Ch.3 <-> Data Pointer/CurrentSetpointValues[2]
//     Term 46 (AT2200-0500)/CC Outputs/Current setpoint value Ch.30 <-> Data Pointer/CurrentSetpointValues[29]
//     Term 46 (AT2200-0500)/CC Outputs/Current setpoint value Ch.4 <-> Data Pointer/CurrentSetpointValues[3]
//     Term 46 (AT2200-0500)/CC Outputs/Current setpoint value Ch.5 <-> Data Pointer/CurrentSetpointValues[4]
//     Term 46 (AT2200-0500)/CC Outputs/Current setpoint value Ch.6 <-> Data Pointer/CurrentSetpointValues[5]
//     Term 46 (AT2200-0500)/CC Outputs/Current setpoint value Ch.7 <-> Data Pointer/CurrentSetpointValues[6]
//     Term 46 (AT2200-0500)/CC Outputs/Current setpoint value Ch.8 <-> Data Pointer/CurrentSetpointValues[7]
//     Term 46 (AT2200-0500)/CC Outputs/Current setpoint value Ch.9 <-> Data Pointer/CurrentSetpointValues[8]
//     Term 46 (AT2200-0500)/LFB Inputs/BinaryData <-> Data Pointer/HallSensorValues
//   Device 40 <-> TcCOM Objects/XTS ProcessingUnit 1/Part 1/Module 54
//     Term 47 (AT2200-0500)/CC Inputs/Current actual value Ch.1 <-> Data Pointer/CurrentActualValues[0]
//     Term 47 (AT2200-0500)/CC Inputs/Current actual value Ch.10 <-> Data Pointer/CurrentActualValues[9]
//     Term 47 (AT2200-0500)/CC Inputs/Current actual value Ch.11 <-> Data Pointer/CurrentActualValues[10]
//     Term 47 (AT2200-0500)/CC Inputs/Current actual value Ch.12 <-> Data Pointer/CurrentActualValues[11]
//     Term 47 (AT2200-0500)/CC Inputs/Current actual value Ch.13 <-> Data Pointer/CurrentActualValues[12]
//     Term 47 (AT2200-0500)/CC Inputs/Current actual value Ch.14 <-> Data Pointer/CurrentActualValues[13]
//     Term 47 (AT2200-0500)/CC Inputs/Current actual value Ch.15 <-> Data Pointer/CurrentActualValues[14]
//     Term 47 (AT2200-0500)/CC Inputs/Current actual value Ch.16 <-> Data Pointer/CurrentActualValues[15]
//     Term 47 (AT2200-0500)/CC Inputs/Current actual value Ch.17 <-> Data Pointer/CurrentActualValues[16]
//     Term 47 (AT2200-0500)/CC Inputs/Current actual value Ch.18 <-> Data Pointer/CurrentActualValues[17]
//     Term 47 (AT2200-0500)/CC Inputs/Current actual value Ch.19 <-> Data Pointer/CurrentActualValues[18]
//     Term 47 (AT2200-0500)/CC Inputs/Current actual value Ch.2 <-> Data Pointer/CurrentActualValues[1]
//     Term 47 (AT2200-0500)/CC Inputs/Current actual value Ch.20 <-> Data Pointer/CurrentActualValues[19]
//     Term 47 (AT2200-0500)/CC Inputs/Current actual value Ch.21 <-> Data Pointer/CurrentActualValues[20]
//     Term 47 (AT2200-0500)/CC Inputs/Current actual value Ch.22 <-> Data Pointer/CurrentActualValues[21]
//     Term 47 (AT2200-0500)/CC Inputs/Current actual value Ch.23 <-> Data Pointer/CurrentActualValues[22]
//     Term 47 (AT2200-0500)/CC Inputs/Current actual value Ch.24 <-> Data Pointer/CurrentActualValues[23]
//     Term 47 (AT2200-0500)/CC Inputs/Current actual value Ch.25 <-> Data Pointer/CurrentActualValues[24]
//     Term 47 (AT2200-0500)/CC Inputs/Current actual value Ch.26 <-> Data Pointer/CurrentActualValues[25]
//     Term 47 (AT2200-0500)/CC Inputs/Current actual value Ch.27 <-> Data Pointer/CurrentActualValues[26]
//     Term 47 (AT2200-0500)/CC Inputs/Current actual value Ch.28 <-> Data Pointer/CurrentActualValues[27]
//     Term 47 (AT2200-0500)/CC Inputs/Current actual value Ch.29 <-> Data Pointer/CurrentActualValues[28]
//     Term 47 (AT2200-0500)/CC Inputs/Current actual value Ch.3 <-> Data Pointer/CurrentActualValues[2]
//     Term 47 (AT2200-0500)/CC Inputs/Current actual value Ch.30 <-> Data Pointer/CurrentActualValues[29]
//     Term 47 (AT2200-0500)/CC Inputs/Current actual value Ch.4 <-> Data Pointer/CurrentActualValues[3]
//     Term 47 (AT2200-0500)/CC Inputs/Current actual value Ch.5 <-> Data Pointer/CurrentActualValues[4]
//     Term 47 (AT2200-0500)/CC Inputs/Current actual value Ch.6 <-> Data Pointer/CurrentActualValues[5]
//     Term 47 (AT2200-0500)/CC Inputs/Current actual value Ch.7 <-> Data Pointer/CurrentActualValues[6]
//     Term 47 (AT2200-0500)/CC Inputs/Current actual value Ch.8 <-> Data Pointer/CurrentActualValues[7]
//     Term 47 (AT2200-0500)/CC Inputs/Current actual value Ch.9 <-> Data Pointer/CurrentActualValues[8]
//     Term 47 (AT2200-0500)/CC Inputs/Status <-> Data Pointer/Status
//     Term 47 (AT2200-0500)/CC Outputs/Control <-> Data Pointer/Control
//     Term 47 (AT2200-0500)/CC Outputs/Current setpoint value Ch.1 <-> Data Pointer/CurrentSetpointValues[0]
//     Term 47 (AT2200-0500)/CC Outputs/Current setpoint value Ch.10 <-> Data Pointer/CurrentSetpointValues[9]
//     Term 47 (AT2200-0500)/CC Outputs/Current setpoint value Ch.11 <-> Data Pointer/CurrentSetpointValues[10]
//     Term 47 (AT2200-0500)/CC Outputs/Current setpoint value Ch.12 <-> Data Pointer/CurrentSetpointValues[11]
//     Term 47 (AT2200-0500)/CC Outputs/Current setpoint value Ch.13 <-> Data Pointer/CurrentSetpointValues[12]
//     Term 47 (AT2200-0500)/CC Outputs/Current setpoint value Ch.14 <-> Data Pointer/CurrentSetpointValues[13]
//     Term 47 (AT2200-0500)/CC Outputs/Current setpoint value Ch.15 <-> Data Pointer/CurrentSetpointValues[14]
//     Term 47 (AT2200-0500)/CC Outputs/Current setpoint value Ch.16 <-> Data Pointer/CurrentSetpointValues[15]
//     Term 47 (AT2200-0500)/CC Outputs/Current setpoint value Ch.17 <-> Data Pointer/CurrentSetpointValues[16]
//     Term 47 (AT2200-0500)/CC Outputs/Current setpoint value Ch.18 <-> Data Pointer/CurrentSetpointValues[17]
//     Term 47 (AT2200-0500)/CC Outputs/Current setpoint value Ch.19 <-> Data Pointer/CurrentSetpointValues[18]
//     Term 47 (AT2200-0500)/CC Outputs/Current setpoint value Ch.2 <-> Data Pointer/CurrentSetpointValues[1]
//     Term 47 (AT2200-0500)/CC Outputs/Current setpoint value Ch.20 <-> Data Pointer/CurrentSetpointValues[19]
//     Term 47 (AT2200-0500)/CC Outputs/Current setpoint value Ch.21 <-> Data Pointer/CurrentSetpointValues[20]
//     Term 47 (AT2200-0500)/CC Outputs/Current setpoint value Ch.22 <-> Data Pointer/CurrentSetpointValues[21]
//     Term 47 (AT2200-0500)/CC Outputs/Current setpoint value Ch.23 <-> Data Pointer/CurrentSetpointValues[22]
//     Term 47 (AT2200-0500)/CC Outputs/Current setpoint value Ch.24 <-> Data Pointer/CurrentSetpointValues[23]
//     Term 47 (AT2200-0500)/CC Outputs/Current setpoint value Ch.25 <-> Data Pointer/CurrentSetpointValues[24]
//     Term 47 (AT2200-0500)/CC Outputs/Current setpoint value Ch.26 <-> Data Pointer/CurrentSetpointValues[25]
//     Term 47 (AT2200-0500)/CC Outputs/Current setpoint value Ch.27 <-> Data Pointer/CurrentSetpointValues[26]
//     Term 47 (AT2200-0500)/CC Outputs/Current setpoint value Ch.28 <-> Data Pointer/CurrentSetpointValues[27]
//     Term 47 (AT2200-0500)/CC Outputs/Current setpoint value Ch.29 <-> Data Pointer/CurrentSetpointValues[28]
//     Term 47 (AT2200-0500)/CC Outputs/Current setpoint value Ch.3 <-> Data Pointer/CurrentSetpointValues[2]
//     Term 47 (AT2200-0500)/CC Outputs/Current setpoint value Ch.30 <-> Data Pointer/CurrentSetpointValues[29]
//     Term 47 (AT2200-0500)/CC Outputs/Current setpoint value Ch.4 <-> Data Pointer/CurrentSetpointValues[3]
//     Term 47 (AT2200-0500)/CC Outputs/Current setpoint value Ch.5 <-> Data Pointer/CurrentSetpointValues[4]
//     Term 47 (AT2200-0500)/CC Outputs/Current setpoint value Ch.6 <-> Data Pointer/CurrentSetpointValues[5]
//     Term 47 (AT2200-0500)/CC Outputs/Current setpoint value Ch.7 <-> Data Pointer/CurrentSetpointValues[6]
//     Term 47 (AT2200-0500)/CC Outputs/Current setpoint value Ch.8 <-> Data Pointer/CurrentSetpointValues[7]
//     Term 47 (AT2200-0500)/CC Outputs/Current setpoint value Ch.9 <-> Data Pointer/CurrentSetpointValues[8]
//     Term 47 (AT2200-0500)/LFB Inputs/BinaryData <-> Data Pointer/HallSensorValues
//   Device 41 <-> TcCOM Objects/XTS ProcessingUnit 1/Part 1/Module 55
//     Term 49 (AT2200-0500)/CC Inputs/Current actual value Ch.1 <-> Data Pointer/CurrentActualValues[0]
//     Term 49 (AT2200-0500)/CC Inputs/Current actual value Ch.10 <-> Data Pointer/CurrentActualValues[9]
//     Term 49 (AT2200-0500)/CC Inputs/Current actual value Ch.11 <-> Data Pointer/CurrentActualValues[10]
//     Term 49 (AT2200-0500)/CC Inputs/Current actual value Ch.12 <-> Data Pointer/CurrentActualValues[11]
//     Term 49 (AT2200-0500)/CC Inputs/Current actual value Ch.13 <-> Data Pointer/CurrentActualValues[12]
//     Term 49 (AT2200-0500)/CC Inputs/Current actual value Ch.14 <-> Data Pointer/CurrentActualValues[13]
//     Term 49 (AT2200-0500)/CC Inputs/Current actual value Ch.15 <-> Data Pointer/CurrentActualValues[14]
//     Term 49 (AT2200-0500)/CC Inputs/Current actual value Ch.16 <-> Data Pointer/CurrentActualValues[15]
//     Term 49 (AT2200-0500)/CC Inputs/Current actual value Ch.17 <-> Data Pointer/CurrentActualValues[16]
//     Term 49 (AT2200-0500)/CC Inputs/Current actual value Ch.18 <-> Data Pointer/CurrentActualValues[17]
//     Term 49 (AT2200-0500)/CC Inputs/Current actual value Ch.19 <-> Data Pointer/CurrentActualValues[18]
//     Term 49 (AT2200-0500)/CC Inputs/Current actual value Ch.2 <-> Data Pointer/CurrentActualValues[1]
//     Term 49 (AT2200-0500)/CC Inputs/Current actual value Ch.20 <-> Data Pointer/CurrentActualValues[19]
//     Term 49 (AT2200-0500)/CC Inputs/Current actual value Ch.21 <-> Data Pointer/CurrentActualValues[20]
//     Term 49 (AT2200-0500)/CC Inputs/Current actual value Ch.22 <-> Data Pointer/CurrentActualValues[21]
//     Term 49 (AT2200-0500)/CC Inputs/Current actual value Ch.23 <-> Data Pointer/CurrentActualValues[22]
//     Term 49 (AT2200-0500)/CC Inputs/Current actual value Ch.24 <-> Data Pointer/CurrentActualValues[23]
//     Term 49 (AT2200-0500)/CC Inputs/Current actual value Ch.25 <-> Data Pointer/CurrentActualValues[24]
//     Term 49 (AT2200-0500)/CC Inputs/Current actual value Ch.26 <-> Data Pointer/CurrentActualValues[25]
//     Term 49 (AT2200-0500)/CC Inputs/Current actual value Ch.27 <-> Data Pointer/CurrentActualValues[26]
//     Term 49 (AT2200-0500)/CC Inputs/Current actual value Ch.28 <-> Data Pointer/CurrentActualValues[27]
//     Term 49 (AT2200-0500)/CC Inputs/Current actual value Ch.29 <-> Data Pointer/CurrentActualValues[28]
//     Term 49 (AT2200-0500)/CC Inputs/Current actual value Ch.3 <-> Data Pointer/CurrentActualValues[2]
//     Term 49 (AT2200-0500)/CC Inputs/Current actual value Ch.30 <-> Data Pointer/CurrentActualValues[29]
//     Term 49 (AT2200-0500)/CC Inputs/Current actual value Ch.4 <-> Data Pointer/CurrentActualValues[3]
//     Term 49 (AT2200-0500)/CC Inputs/Current actual value Ch.5 <-> Data Pointer/CurrentActualValues[4]
//     Term 49 (AT2200-0500)/CC Inputs/Current actual value Ch.6 <-> Data Pointer/CurrentActualValues[5]
//     Term 49 (AT2200-0500)/CC Inputs/Current actual value Ch.7 <-> Data Pointer/CurrentActualValues[6]
//     Term 49 (AT2200-0500)/CC Inputs/Current actual value Ch.8 <-> Data Pointer/CurrentActualValues[7]
//     Term 49 (AT2200-0500)/CC Inputs/Current actual value Ch.9 <-> Data Pointer/CurrentActualValues[8]
//     Term 49 (AT2200-0500)/CC Inputs/Status <-> Data Pointer/Status
//     Term 49 (AT2200-0500)/CC Outputs/Control <-> Data Pointer/Control
//     Term 49 (AT2200-0500)/CC Outputs/Current setpoint value Ch.1 <-> Data Pointer/CurrentSetpointValues[0]
//     Term 49 (AT2200-0500)/CC Outputs/Current setpoint value Ch.10 <-> Data Pointer/CurrentSetpointValues[9]
//     Term 49 (AT2200-0500)/CC Outputs/Current setpoint value Ch.11 <-> Data Pointer/CurrentSetpointValues[10]
//     Term 49 (AT2200-0500)/CC Outputs/Current setpoint value Ch.12 <-> Data Pointer/CurrentSetpointValues[11]
//     Term 49 (AT2200-0500)/CC Outputs/Current setpoint value Ch.13 <-> Data Pointer/CurrentSetpointValues[12]
//     Term 49 (AT2200-0500)/CC Outputs/Current setpoint value Ch.14 <-> Data Pointer/CurrentSetpointValues[13]
//     Term 49 (AT2200-0500)/CC Outputs/Current setpoint value Ch.15 <-> Data Pointer/CurrentSetpointValues[14]
//     Term 49 (AT2200-0500)/CC Outputs/Current setpoint value Ch.16 <-> Data Pointer/CurrentSetpointValues[15]
//     Term 49 (AT2200-0500)/CC Outputs/Current setpoint value Ch.17 <-> Data Pointer/CurrentSetpointValues[16]
//     Term 49 (AT2200-0500)/CC Outputs/Current setpoint value Ch.18 <-> Data Pointer/CurrentSetpointValues[17]
//     Term 49 (AT2200-0500)/CC Outputs/Current setpoint value Ch.19 <-> Data Pointer/CurrentSetpointValues[18]
//     Term 49 (AT2200-0500)/CC Outputs/Current setpoint value Ch.2 <-> Data Pointer/CurrentSetpointValues[1]
//     Term 49 (AT2200-0500)/CC Outputs/Current setpoint value Ch.20 <-> Data Pointer/CurrentSetpointValues[19]
//     Term 49 (AT2200-0500)/CC Outputs/Current setpoint value Ch.21 <-> Data Pointer/CurrentSetpointValues[20]
//     Term 49 (AT2200-0500)/CC Outputs/Current setpoint value Ch.22 <-> Data Pointer/CurrentSetpointValues[21]
//     Term 49 (AT2200-0500)/CC Outputs/Current setpoint value Ch.23 <-> Data Pointer/CurrentSetpointValues[22]
//     Term 49 (AT2200-0500)/CC Outputs/Current setpoint value Ch.24 <-> Data Pointer/CurrentSetpointValues[23]
//     Term 49 (AT2200-0500)/CC Outputs/Current setpoint value Ch.25 <-> Data Pointer/CurrentSetpointValues[24]
//     Term 49 (AT2200-0500)/CC Outputs/Current setpoint value Ch.26 <-> Data Pointer/CurrentSetpointValues[25]
//     Term 49 (AT2200-0500)/CC Outputs/Current setpoint value Ch.27 <-> Data Pointer/CurrentSetpointValues[26]
//     Term 49 (AT2200-0500)/CC Outputs/Current setpoint value Ch.28 <-> Data Pointer/CurrentSetpointValues[27]
//     Term 49 (AT2200-0500)/CC Outputs/Current setpoint value Ch.29 <-> Data Pointer/CurrentSetpointValues[28]
//     Term 49 (AT2200-0500)/CC Outputs/Current setpoint value Ch.3 <-> Data Pointer/CurrentSetpointValues[2]
